   #r := FALSE;
   #a1 := W#16#0000;
   #a2 := W#16#0000;
   #activeDataBlock := 0;
   // PB17, STEP 5 network 1
   #r := ((NOT "ROLL_State".M[70, 1]) AND "ROLL_State".M[3, 3]);
   "ROLL_State".M[70, 0] := #r;
   // PB17, STEP 5 network 2
   #r := "ROLL_State".M[70, 0];
   IF #r THEN
       "ROLL_State".M[70, 1] := TRUE;
   END_IF;
   #r := "ROLL_IO".Input[0, 2];
   IF #r THEN
       "ROLL_State".M[70, 1] := FALSE;
   END_IF;
   // PB17, STEP 5 network 3
   #r := ((("ROLL_IO".Input[0, 1] AND "ROLL_State".M[74, 1]) OR ("ROLL_IO".Input[0, 2] AND "ROLL_State".M[64, 0])) AND "ROLL_State".M[29, 1]);
   "ROLL_IO".Output[112, 0] := #r;
   // PB17, STEP 5 network 4
   #r := ((("ROLL_IO".Input[0, 1] AND "ROLL_State".M[74, 5]) OR ("ROLL_IO".Input[0, 2] AND "ROLL_State".M[64, 1])) AND "ROLL_State".M[29, 1]);
   "ROLL_IO".Output[112, 5] := #r;
   // PB17, STEP 5 network 5
   #r := (((("ROLL_IO".Input[0, 1] AND "ROLL_State".M[78, 4]) OR ("ROLL_IO".Input[0, 2] AND "ROLL_State".M[64, 4])) AND "ROLL_State".M[29, 0]) OR ("ROLL_IO".Output[113, 1] AND "ROLL_IO".Output[113, 3]));
   "ROLL_IO".Output[113, 1] := #r;
   // PB17, STEP 5 network 6
   #r := (((NOT "ROLL_State".M[71, 4]) AND "ROLL_State".M[71, 3]) OR ((("ROLL_IO".Input[0, 1] AND "ROLL_State".M[78, 6]) OR ("ROLL_IO".Input[0, 2] AND "ROLL_State".M[64, 5])) AND "ROLL_State".M[29, 0]));
   "ROLL_State".M[71, 3] := #r;
   // PB17, STEP 5 network 7
   #r := "ROLL_State".M[71, 3];
   "ROLL_IO".Output[113, 3] := #r;
   // PB17, STEP 5 network 8
   #r := (((NOT "ROLL_State".M[71, 3]) AND "ROLL_State".M[71, 4]) OR ((((NOT "ROLL_State".M[64, 5]) AND ((NOT "ROLL_State".M[20, 2]) OR "ROLL_IO".Input[124, 5]) AND "ROLL_IO".Input[0, 2]) OR ("ROLL_IO".Input[0, 1] AND "ROLL_State".M[78, 7])) AND "ROLL_State".M[29, 0]));
   "ROLL_State".M[71, 4] := #r;
   // PB17, STEP 5 network 9
   #r := "ROLL_State".M[71, 4];
   "ROLL_IO".Output[113, 2] := #r;
   // PB17, STEP 5 network 10
   #r := (("ROLL_IO".Input[0, 1] AND "ROLL_State".M[75, 4]) OR ("ROLL_IO".Input[0, 2] AND "ROLL_State".M[35, 2] AND "ROLL_State".M[65, 0]));
   "ROLL_State".M[79, 5] := #r;
   // PB17, STEP 5 network 11
   #r := ((NOT "ROLL_IO".Output[23, 0]) AND (NOT "ROLL_IO".Output[23, 4]) AND (NOT "ROLL_State".M[10, 3]) AND (NOT "ROLL_State".M[5, 0]) AND ((NOT "ROLL_IO".Input[11, 4]) OR (NOT "ROLL_IO".Input[11, 6])) AND "ROLL_IO".Input[11, 7] AND "ROLL_IO".Input[12, 5] AND "ROLL_IO".Input[12, 7] AND "ROLL_IO".Input[14, 0] AND "ROLL_State".M[29, 0] AND "ROLL_State".M[79, 5]);
   "ROLL_IO".Output[23, 1] := #r;
   // PB17, STEP 5 network 12
   #r := (("ROLL_IO".Input[0, 1] AND "ROLL_State".M[75, 5]) OR ("ROLL_IO".Input[0, 2] AND "ROLL_State".M[35, 2] AND "ROLL_State".M[65, 5]));
   "ROLL_State".M[79, 6] := #r;
   // PB17, STEP 5 network 13
   #r := ((NOT "ROLL_IO".Output[23, 1]) AND (NOT "ROLL_IO".Output[23, 4]) AND (NOT "ROLL_State".M[10, 2]) AND (NOT "ROLL_State".M[5, 0]) AND (((NOT "ROLL_IO".Input[119, 0]) AND "ROLL_State".M[0, 3]) OR (NOT "ROLL_IO".Input[11, 0]) OR (NOT "ROLL_IO".Input[11, 6])) AND "ROLL_IO".Input[11, 7] AND "ROLL_IO".Input[12, 5] AND "ROLL_IO".Input[12, 7] AND "ROLL_IO".Input[14, 0] AND "ROLL_State".M[29, 0] AND "ROLL_State".M[79, 6]);
   "ROLL_IO".Output[23, 0] := #r;
   // PB17, STEP 5 network 14
   #r := ((("ROLL_IO".Input[0, 1] AND "ROLL_State".M[75, 6]) OR ("ROLL_IO".Input[0, 2] AND "ROLL_State".M[35, 2] AND "ROLL_State".M[65, 6])) AND ("ROLL_IO".Output[23, 0] OR "ROLL_IO".Output[23, 1]));
   "ROLL_IO".Output[23, 3] := #r;
   // PB17, STEP 5 network 15
   #r := ((NOT "ROLL_IO".Output[23, 3]) AND ("ROLL_IO".Output[23, 0] OR "ROLL_IO".Output[23, 1]) AND ("ROLL_IO".Input[0, 1] OR "ROLL_State".M[31, 5]) AND "ROLL_State".M[29, 0]);
   "ROLL_IO".Output[23, 2] := #r;
   // PB17, STEP 5 network 16
   #r := (("ROLL_IO".Input[0, 1] AND "ROLL_State".M[76, 2]) OR ("ROLL_IO".Input[0, 2] AND "ROLL_State".M[35, 2] AND "ROLL_State".M[66, 4]));
   "ROLL_State".M[80, 0] := #r;
   // PB17, STEP 5 network 17
   #r := ((NOT "ROLL_IO".Output[23, 4]) AND (NOT "ROLL_State".M[10, 1]) AND (NOT "ROLL_State".M[5, 2]) AND (NOT "ROLL_State".M[9, 0]) AND ((NOT "ROLL_IO".Input[12, 5]) OR (NOT "ROLL_IO".Input[12, 7])) AND ("ROLL_IO".Input[124, 2] OR "ROLL_State".M[0, 4]) AND "ROLL_IO".Input[13, 0] AND "ROLL_IO".Input[13, 7] AND "ROLL_IO".Input[14, 0] AND "ROLL_State".M[29, 0] AND "ROLL_State".M[80, 0]);
   "ROLL_IO".Output[23, 5] := #r;
   // PB17, STEP 5 network 18
   #r := (("ROLL_IO".Input[0, 1] AND "ROLL_State".M[77, 0]) OR ("ROLL_IO".Input[0, 2] AND "ROLL_State".M[35, 2] AND "ROLL_State".M[66, 7]));
   "ROLL_State".M[80, 1] := #r;
   // PB17, STEP 5 network 19
   #r := "ROLL_IO".Input[12, 5];
   IF #r THEN
       "ROLL_State".M[80, 2] := TRUE;
   END_IF;
   #r := "ROLL_IO".Input[12, 1];
   IF #r THEN
       "ROLL_State".M[80, 2] := FALSE;
   END_IF;
   // PB17, STEP 5 network 20
   #r := (((("ROLL_IO".Input[11, 1] OR "ROLL_IO".Input[11, 2] OR "ROLL_IO".Input[11, 3] OR "ROLL_IO".Input[11, 4] OR "ROLL_IO".Input[119, 6] OR "ROLL_IO".Input[119, 7] OR "ROLL_IO".Input[120, 0] OR "ROLL_IO".Input[120, 1]) AND "ROLL_IO".Input[12, 1]) OR ("ROLL_IO".Input[11, 0] AND "ROLL_IO".Input[12, 1])) AND "ROLL_IO".Input[12, 7]);
   "ROLL_State".M[80, 6] := #r;
   // PB17, STEP 5 network 21
   #r := (("ROLL_IO".Input[11, 0] OR "ROLL_IO".Input[11, 1] OR "ROLL_IO".Input[11, 2] OR "ROLL_IO".Input[11, 3] OR "ROLL_IO".Input[11, 4] OR "ROLL_IO".Input[119, 6] OR "ROLL_IO".Input[119, 7] OR "ROLL_IO".Input[120, 0] OR "ROLL_IO".Input[120, 1]) AND "ROLL_IO".Input[12, 5] AND "ROLL_IO".Input[12, 7]);
   "ROLL_State".M[80, 7] := #r;
   // PB17, STEP 5 network 22
   #r := ((NOT "ROLL_IO".Output[23, 0]) AND (NOT "ROLL_IO".Output[23, 1]) AND (NOT "ROLL_IO".Output[23, 5]) AND (NOT "ROLL_State".M[10, 0]) AND (NOT "ROLL_State".M[5, 2]) AND (NOT "ROLL_State".M[80, 6]) AND ("ROLL_IO".Input[124, 2] OR "ROLL_State".M[0, 4]) AND "ROLL_IO".Input[13, 0] AND "ROLL_IO".Input[14, 0] AND "ROLL_State".M[29, 0] AND "ROLL_State".M[80, 1]);
   "ROLL_IO".Output[23, 4] := #r;
   // PB17, STEP 5 network 23
   #r := ((NOT "ROLL_State".M[68, 2]) AND (((NOT "ROLL_IO".Input[12, 5]) AND "ROLL_IO".Output[23, 5]) OR ("ROLL_IO".Output[23, 4] AND "ROLL_State".M[80, 2])));
   "ROLL_IO".Output[23, 7] := #r;
   // PB17, STEP 5 network 24
   #r := ((NOT "ROLL_IO".Output[23, 7]) AND ("ROLL_IO".Output[23, 4] OR "ROLL_IO".Output[23, 5]));
   "ROLL_IO".Output[23, 6] := #r;
   // PB17, STEP 5 network 25
   #r := (("ROLL_IO".Input[0, 1] AND "ROLL_State".M[77, 6]) OR ("ROLL_IO".Input[0, 2] AND "ROLL_State".M[35, 2] AND "ROLL_State".M[67, 0]));
   "ROLL_State".M[80, 3] := #r;
   // PB17, STEP 5 network 26
   #r := ((NOT "ROLL_IO".Output[112, 1]) AND (NOT "ROLL_IO".Output[113, 3]) AND (NOT "ROLL_IO".Input[124, 2]) AND (NOT "ROLL_State".M[10, 5]) AND (NOT "ROLL_State".M[70, 2]) AND (NOT "ROLL_State".M[9, 3]) AND "ROLL_IO".Input[11, 0] AND "ROLL_IO".Input[11, 6] AND "ROLL_IO".Input[12, 1] AND "ROLL_IO".Input[12, 7] AND "ROLL_State".M[29, 0] AND "ROLL_State".M[80, 3]);
   "ROLL_IO".Output[112, 2] := #r;
   // PB17, STEP 5 network 27
   #r := (("ROLL_IO".Input[0, 1] AND "ROLL_State".M[77, 4]) OR ("ROLL_IO".Input[0, 2] AND "ROLL_State".M[35, 2] AND "ROLL_State".M[67, 1]));
   "ROLL_State".M[80, 4] := #r;
   // PB17, STEP 5 network 28
   #r := ((NOT "ROLL_IO".Output[112, 2]) AND (NOT "ROLL_IO".Output[113, 3]) AND (NOT "ROLL_IO".Input[124, 1]) AND (NOT "ROLL_State".M[10, 4]) AND (NOT "ROLL_State".M[70, 2]) AND (NOT "ROLL_State".M[70, 3]) AND (NOT "ROLL_State".M[9, 3]) AND "ROLL_IO".Input[11, 0] AND "ROLL_IO".Input[11, 6] AND "ROLL_IO".Input[12, 1] AND "ROLL_IO".Input[12, 7] AND "ROLL_State".M[29, 0] AND "ROLL_State".M[80, 4]);
   "ROLL_IO".Output[112, 1] := #r;
   // PB17, STEP 5 network 29
   #r := ((("ROLL_IO".Input[0, 1] AND "ROLL_State".M[77, 7]) OR ("ROLL_IO".Input[0, 2] AND "ROLL_State".M[35, 2] AND "ROLL_State".M[67, 5])) AND "ROLL_State".M[29, 0]);
   "ROLL_IO".Output[112, 4] := #r;
   // PB17, STEP 5 network 30
   #r := ((("ROLL_IO".Input[0, 1] AND "ROLL_State".M[78, 0]) OR ("ROLL_IO".Input[0, 2] AND "ROLL_State".M[35, 2] AND "ROLL_State".M[67, 6])) AND "ROLL_State".M[29, 0]);
   "ROLL_IO".Output[112, 3] := #r;
   // PB17, STEP 5 network 31
   #r := ((NOT "ROLL_State".M[16, 0]) AND (NOT "ROLL_State".M[16, 1]) AND (NOT "ROLL_State".M[16, 2]) AND (NOT "ROLL_State".M[16, 4]) AND "ROLL_State".M[37, 2]);
   "ROLL_State".M[81, 4] := #r;
   // PB17, STEP 5 network 32
   RETURN;
END_FUNCTION

FUNCTION "ROLL_PB18" : Void   // FC26, SCL
{ S7_Optimized_Access := 'TRUE' }
VERSION : 0.1
// stored: AutoNumber true, IsIECCheckEnabled false, SetENOAutomatically false, UDAEnableTagReadback false
   VAR_TEMP
      r : Bool;
      a1 : Word;
      a2 : Word;
      activeDataBlock : Int;
      comparisonResults : Array[0..0] of Bool;
   END_VAR
BEGIN

   #r := FALSE;
   #a1 := W#16#0000;
   #a2 := W#16#0000;
   #activeDataBlock := 0;
   // PB18, STEP 5 network 1
   #r := ("ROLL_State".M[70, 2] OR "ROLL_State".M[70, 3] OR "ROLL_State".M[70, 4] OR "ROLL_State".M[70, 6] OR "ROLL_State".M[71, 0]);
   "ROLL_State".M[80, 5] := #r;
   // PB18, STEP 5 network 2
   #r := (((NOT "ROLL_IO".Output[112, 0]) AND (NOT "ROLL_IO".Output[112, 5]) AND "ROLL_State".M[20, 5]) OR ((NOT "ROLL_IO".Output[112, 0]) AND "ROLL_State".M[20, 3]) OR ((NOT "ROLL_IO".Output[112, 5]) AND "ROLL_State".M[20, 4]) OR ((NOT "ROLL_IO".Output[17, 7]) AND "ROLL_State".M[20, 7]) OR (("ROLL_State".M[20, 1] OR "ROLL_State".M[20, 2]) AND "ROLL_State".M[28, 4]));
   "ROLL_State".M[250, 0] := #r;
   // PB18, STEP 5 network 3
   #r := (((NOT "ROLL_IO".Output[113, 0]) AND "ROLL_State".M[22, 2]) OR ((NOT "ROLL_IO".Output[113, 1]) AND "ROLL_State".M[22, 3]) OR ((NOT "ROLL_IO".Output[113, 3]) AND "ROLL_IO".Output[113, 2] AND "ROLL_State".M[22, 4]) OR ((NOT "ROLL_IO".Output[113, 5]) AND "ROLL_IO".Output[113, 4] AND "ROLL_State".M[22, 5]) OR ("ROLL_IO".Input[124, 1] AND "ROLL_State".M[22, 0]) OR ("ROLL_IO".Input[124, 4] AND "ROLL_State".M[22, 1]) OR "ROLL_State".M[250, 0]);
   "ROLL_State".M[250, 0] := #r;
   // PB18, STEP 5 network 4
   #r := ((("ROLL_IO".Input[11, 1] OR "ROLL_IO".Input[11, 2] OR "ROLL_IO".Input[11, 3] OR "ROLL_IO".Input[11, 4] OR "ROLL_IO".Input[119, 6] OR "ROLL_IO".Input[119, 7] OR "ROLL_IO".Input[120, 0] OR "ROLL_IO".Input[120, 1]) AND "ROLL_IO".Input[12, 5] AND "ROLL_IO".Input[12, 7] AND "ROLL_State".M[23, 0]) OR (("ROLL_State".M[23, 2] OR "ROLL_State".M[23, 3]) AND "ROLL_State".M[63, 1]) OR ("ROLL_IO".Input[11, 0] AND "ROLL_IO".Input[11, 6] AND "ROLL_State".M[23, 1]) OR ("ROLL_IO".Input[11, 0] AND "ROLL_IO".Input[12, 1] AND "ROLL_IO".Input[12, 7] AND "ROLL_State".M[23, 0]) OR "ROLL_State".M[250, 0]);
   "ROLL_State".M[250, 0] := #r;
   // PB18, STEP 5 network 5
   #r := (((NOT "ROLL_IO".Output[20, 1]) AND "ROLL_State".M[24, 1]) OR "ROLL_State".M[250, 0]);
   "ROLL_State".M[250, 0] := #r;
   // PB18, STEP 5 network 6
   #r := ((((NOT "ROLL_IO".Output[20, 4]) OR (NOT "ROLL_IO".Output[22, 6])) AND "ROLL_State".M[25, 0]) OR "ROLL_State".M[250, 0]);
   "ROLL_State".M[250, 0] := #r;
   // PB18, STEP 5 network 7
   #r := (((NOT "ROLL_IO".Output[20, 5]) AND "ROLL_State".M[26, 6]) OR ((NOT "ROLL_IO".Output[20, 6]) AND "ROLL_State".M[26, 0]) OR ((NOT "ROLL_IO".Output[21, 4]) AND "ROLL_State".M[26, 5]) OR "ROLL_State".M[250, 0]);
   "ROLL_State".M[250, 0] := #r;
   // PB18, STEP 5 network 8
   #r := (((NOT "ROLL_IO".Output[20, 6]) AND "ROLL_State".M[27, 4]) OR ((NOT "ROLL_IO".Output[21, 6]) AND "ROLL_State".M[27, 5]) OR ((NOT "ROLL_State".M[80, 5]) AND "ROLL_State".M[27, 7]) OR "ROLL_State".M[250, 0]);
   "ROLL_State".M[250, 0] := #r;
   // PB18, STEP 5 network 9
   #r := ((("ROLL_IO".Output[112, 0] OR "ROLL_IO".Output[112, 5]) AND "ROLL_State".M[20, 5]) OR ("ROLL_IO".Output[112, 0] AND "ROLL_State".M[20, 3]) OR ("ROLL_IO".Output[112, 5] AND "ROLL_State".M[20, 4]) OR ("ROLL_IO".Output[17, 7] AND "ROLL_State".M[20, 7]));
   "ROLL_State".M[252, 0] := #r;
   // PB18, STEP 5 network 10
   #r := (((NOT "ROLL_IO".Output[113, 2]) AND "ROLL_IO".Output[113, 3] AND "ROLL_State".M[22, 4]) OR ((NOT "ROLL_IO".Output[113, 4]) AND "ROLL_IO".Output[113, 5] AND "ROLL_State".M[22, 5]) OR ("ROLL_IO".Output[113, 0] AND "ROLL_State".M[22, 2]) OR ("ROLL_IO".Output[113, 1] AND "ROLL_State".M[22, 3]) OR ("ROLL_IO".Input[124, 2] AND "ROLL_State".M[22, 0]) OR ("ROLL_IO".Input[124, 5] AND "ROLL_State".M[22, 1]) OR "ROLL_State".M[252, 0]);
   "ROLL_State".M[252, 0] := #r;
   // PB18, STEP 5 network 11
   #r := (((NOT "ROLL_IO".Output[23, 1]) AND ("ROLL_IO".Input[11, 1] OR "ROLL_IO".Input[11, 2] OR "ROLL_IO".Input[11, 3] OR "ROLL_IO".Input[11, 4] OR "ROLL_IO".Input[119, 6] OR "ROLL_IO".Input[119, 7] OR "ROLL_IO".Input[120, 0] OR "ROLL_IO".Input[120, 1]) AND "ROLL_IO".Input[11, 6] AND "ROLL_State".M[23, 1]) OR ((NOT "ROLL_State".M[63, 1]) AND ("ROLL_State".M[23, 2] OR "ROLL_State".M[23, 3])) OR (((("ROLL_IO".Input[11, 1] OR "ROLL_IO".Input[11, 2] OR "ROLL_IO".Input[11, 3] OR "ROLL_IO".Input[11, 4] OR "ROLL_IO".Input[119, 6] OR "ROLL_IO".Input[119, 7] OR "ROLL_IO".Input[120, 0] OR "ROLL_IO".Input[120, 1]) AND "ROLL_IO".Input[12, 1]) OR ("ROLL_IO".Input[11, 0] AND "ROLL_IO".Input[12, 5])) AND "ROLL_IO".Input[12, 7] AND "ROLL_State".M[23, 0]) OR "ROLL_State".M[252, 0]);
   "ROLL_State".M[252, 0] := #r;
   // PB18, STEP 5 network 12
   #r := (("ROLL_IO".Output[20, 1] AND "ROLL_State".M[24, 1]) OR "ROLL_State".M[252, 0]);
   "ROLL_State".M[252, 0] := #r;
   // PB18, STEP 5 network 13
   #r := (("ROLL_IO".Output[20, 4] AND "ROLL_IO".Output[22, 6] AND "ROLL_State".M[25, 0]) OR "ROLL_State".M[252, 0]);
   "ROLL_State".M[252, 0] := #r;
   // PB18, STEP 5 network 14
   #r := (("ROLL_IO".Output[20, 6] AND "ROLL_State".M[26, 0]) OR "ROLL_State".M[252, 0]);
   "ROLL_State".M[252, 0] := #r;
   // PB18, STEP 5 network 15
   #r := (("ROLL_IO".Output[20, 5] AND "ROLL_State".M[26, 6]) OR ("ROLL_IO".Output[20, 6] AND "ROLL_State".M[27, 4]) OR ("ROLL_IO".Output[21, 4] AND "ROLL_State".M[26, 5]) OR ("ROLL_IO".Output[21, 6] AND "ROLL_State".M[27, 5]) OR ("ROLL_State".M[27, 7] AND "ROLL_State".M[80, 5]) OR "ROLL_State".M[252, 0]);
   "ROLL_State".M[252, 0] := #r;
   // PB18, STEP 5 network 16
   RETURN;
END_FUNCTION

FUNCTION "ROLL_PB19" : Void   // FC27, SCL
{ S7_Optimized_Access := 'TRUE' }
VERSION : 0.1
// stored: AutoNumber true, IsIECCheckEnabled false, SetENOAutomatically false, UDAEnableTagReadback false
   VAR_TEMP
      r : Bool;
      a1 : Word;
      a2 : Word;
      activeDataBlock : Int;
      comparisonResults : Array[0..0] of Bool;
   END_VAR
BEGIN

   #r := FALSE;
   #a1 := W#16#0000;
   #a2 := W#16#0000;
   #activeDataBlock := 0;
   // PB19, STEP 5 network 1
   #r := ((NOT "ROLL_IO".Input[3, 6]) AND (NOT "ROLL_State".M[5, 6]) AND (NOT "ROLL_State".M[6, 0]) AND (NOT "ROLL_State".M[6, 2]) AND ("ROLL_IO".Input[3, 1] OR "ROLL_State".M[31, 5]) AND "ROLL_IO".Input[5, 2] AND "ROLL_IO".Input[5, 4] AND "ROLL_State".M[4, 1]);
   "ROLL_State".M[82, 0] := #r;
   // PB19, STEP 5 network 2
   #r := ((NOT "ROLL_IO".Input[3, 6]) AND (NOT "ROLL_State".M[12, 0]) AND (NOT "ROLL_State".M[5, 3]) AND (NOT "ROLL_State".M[5, 6]) AND ("ROLL_IO".Input[3, 1] OR "ROLL_State".M[31, 5]) AND "ROLL_IO".Input[8, 3] AND "ROLL_IO".Input[8, 5] AND "ROLL_State".M[4, 1]);
   "ROLL_State".M[82, 2] := #r;
   // PB19, STEP 5 network 3
   #r := ("ROLL_State".M[31, 5] AND "ROLL_State".M[40, 0]);
   IF #r THEN
       "ROLL_State".M[82, 3] := TRUE;
   END_IF;
   #r := (NOT "ROLL_State".M[31, 5]);
   IF #r THEN
       "ROLL_State".M[82, 3] := FALSE;
   END_IF;
   // PB19, STEP 5 network 4
   #r := ((NOT "ROLL_State".M[110, 1]) AND (NOT "ROLL_State".M[110, 2]) AND "ROLL_State".M[110, 0] AND "ROLL_State".M[110, 3] AND "ROLL_State".M[40, 0]);
   "ROLL_State".M[240, 0] := #r;
   // PB19, STEP 5 network 5
   #r := (((NOT "ROLL_State".M[110, 2]) AND "ROLL_State".M[110, 0] AND "ROLL_State".M[110, 1] AND "ROLL_State".M[110, 3] AND "ROLL_State".M[41, 1]) OR "ROLL_State".M[240, 0]);
   "ROLL_State".M[240, 0] := #r;
   // PB19, STEP 5 network 6
   #r := (((NOT "ROLL_State".M[110, 1]) AND "ROLL_State".M[110, 0] AND "ROLL_State".M[110, 2] AND "ROLL_State".M[110, 3] AND "ROLL_State".M[41, 1]) OR "ROLL_State".M[240, 0]);
   "ROLL_State".M[240, 0] := #r;
   // PB19, STEP 5 network 7
   #r := (("ROLL_State".M[110, 0] AND "ROLL_State".M[110, 1] AND "ROLL_State".M[110, 2] AND "ROLL_State".M[110, 3] AND "ROLL_State".M[41, 1]) OR "ROLL_State".M[240, 0]);
   "ROLL_State".M[240, 0] := #r;
   // PB19, STEP 5 network 8
   #r := ("ROLL_State".M[240, 0] AND "ROLL_State".M[31, 5]);
   IF #r THEN
       "ROLL_State".M[82, 4] := TRUE;
   END_IF;
   #r := ((NOT "ROLL_State".M[31, 5]) OR "ROLL_State".M[45, 5]);
   IF #r THEN
       "ROLL_State".M[82, 4] := FALSE;
   END_IF;
   // PB19, STEP 5 network 9
   #r := ((NOT "ROLL_IO".Output[17, 3]) AND (NOT "ROLL_State".M[82, 4]) AND (NOT "ROLL_State".S5Timers[91].Q) AND ("ROLL_State".M[82, 3] OR "ROLL_State".S5Timers[22].Q) AND "ROLL_IO".Input[8, 5]);
   "ROLL_IO".Output[17, 2] := #r;
   // PB19, STEP 5 network 10
   #r := ((NOT "ROLL_IO".Output[17, 2]) AND (NOT "ROLL_State".S5Timers[90].Q) AND "ROLL_IO".Input[3, 0] AND "ROLL_IO".Input[8, 5] AND "ROLL_State".M[82, 4]);
   "ROLL_IO".Output[17, 3] := #r;
   // PB19, STEP 5 network 11
   #a2 := #a1;
   #a1 := W#16#3060;
   #r := "ROLL_IO".Output[18, 0];
   "ROLL_TimerOp"(Number := 22,
                  Operation := 1,
                  Signal := #r,
                  Preset := #a1);
   // PB19, STEP 5 network 12
   #a2 := #a1;
   #a1 := W#16#1005;
   #r := "ROLL_IO".Output[17, 2];
   "ROLL_TimerOp"(Number := 90,
                  Operation := 1,
                  Signal := #r,
                  Preset := #a1);
   // PB19, STEP 5 network 13
   #a2 := #a1;
   #a1 := W#16#1040;
   #r := "ROLL_IO".Output[17, 3];
   "ROLL_TimerOp"(Number := 91,
                  Operation := 1,
                  Signal := #r,
                  Preset := #a1);
   // PB19, STEP 5 network 14
   #r := ((NOT "ROLL_State".M[12, 0]) AND (NOT "ROLL_State".M[19, 7]) AND ("ROLL_IO".Output[17, 2] OR "ROLL_IO".Output[17, 3] OR "ROLL_State".S5Timers[90].Q OR "ROLL_State".S5Timers[91].Q) AND ("ROLL_State".M[82, 3] OR "ROLL_State".M[82, 4]) AND "ROLL_IO".Input[8, 3] AND "ROLL_IO".Input[8, 4] AND "ROLL_State".M[82, 2]);
   "ROLL_IO".Output[18, 0] := #r;
   // PB19, STEP 5 network 15
   #r := "ROLL_IO".Output[18, 0];
   "ROLL_IO".Output[18, 1] := #r;
   // PB19, STEP 5 network 16
   #r := ("ROLL_IO".Output[18, 0] AND "ROLL_State".M[82, 4]);
   "ROLL_IO".Output[18, 2] := #r;
   // PB19, STEP 5 network 17
   #r := ("ROLL_IO".Output[18, 0] AND "ROLL_State".M[82, 4]);
   "ROLL_IO".Output[18, 3] := #r;
   // PB19, STEP 5 network 18
   RETURN;
END_FUNCTION

FUNCTION "ROLL_PB2" : Void   // FC14, SCL
{ S7_Optimized_Access := 'TRUE' }
VERSION : 0.1
// stored: AutoNumber true, IsIECCheckEnabled false, SetENOAutomatically false, UDAEnableTagReadback false
   VAR_TEMP
      r : Bool;
      a1 : Word;
      a2 : Word;
      activeDataBlock : Int;
      comparisonResults : Array[0..0] of Bool;
   END_VAR
BEGIN

   #r := FALSE;
   #a1 := W#16#0000;
   #a2 := W#16#0000;
   #activeDataBlock := 0;
   // PB2, STEP 5 network 1
   #r := ((NOT "ROLL_State".M[0, 1]) AND "ROLL_State".S5Timers[11].Q);
   "ROLL_State".M[4, 1] := #r;
   // PB2, STEP 5 network 2
   #r := ((NOT "ROLL_State".M[4, 1]) OR "ROLL_IO".Input[1, 0]);
   "ROLL_State".M[3, 1] := #r;
   // PB2, STEP 5 network 3
   #r := ((((NOT "ROLL_State".M[31, 4]) AND "ROLL_IO".Input[0, 4] AND "ROLL_State".M[4, 1]) OR "ROLL_State".M[31, 5]) AND "ROLL_IO".Input[0, 2]);
   "ROLL_State".M[4, 4] := #r;
   // PB2, STEP 5 network 4
   #r := (NOT "ROLL_IO".Input[11, 7]);
   IF #r THEN
       "ROLL_State".M[5, 0] := TRUE;
   END_IF;
   #r := "ROLL_State".M[3, 1];
   IF #r THEN
       "ROLL_State".M[5, 0] := FALSE;
   END_IF;
   // PB2, STEP 5 network 5
   #r := (NOT "ROLL_IO".Input[13, 5]);
   IF #r THEN
       "ROLL_State".M[5, 1] := TRUE;
   END_IF;
   #r := "ROLL_State".M[3, 1];
   IF #r THEN
       "ROLL_State".M[5, 1] := FALSE;
   END_IF;
   // PB2, STEP 5 network 6
   #r := (NOT "ROLL_IO".Input[13, 0]);
   IF #r THEN
       "ROLL_State".M[5, 2] := TRUE;
   END_IF;
   #r := "ROLL_State".M[3, 1];
   IF #r THEN
       "ROLL_State".M[5, 2] := FALSE;
   END_IF;
   // PB2, STEP 5 network 7
   #r := (NOT "ROLL_IO".Input[8, 5]);
   IF #r THEN
       "ROLL_State".M[5, 3] := TRUE;
   END_IF;
   #r := "ROLL_State".M[3, 1];
   IF #r THEN
       "ROLL_State".M[5, 3] := FALSE;
   END_IF;
   // PB2, STEP 5 network 8
   #r := "ROLL_State".M[0, 3];
   IF #r THEN
       "ROLL_State".M[5, 4] := TRUE;
   END_IF;
   #r := "ROLL_State".M[3, 1];
   IF #r THEN
       "ROLL_State".M[5, 4] := FALSE;
   END_IF;
   // PB2, STEP 5 network 9
   #r := "ROLL_State".M[0, 3];
   IF #r THEN
       "ROLL_State".M[5, 5] := TRUE;
   END_IF;
   #r := "ROLL_State".M[3, 1];
   IF #r THEN
       "ROLL_State".M[5, 5] := FALSE;
   END_IF;
   // PB2, STEP 5 network 10
   #r := "ROLL_IO".Input[3, 6];
   IF #r THEN
       "ROLL_State".M[5, 6] := TRUE;
   END_IF;
   #r := "ROLL_State".M[3, 1];
   IF #r THEN
       "ROLL_State".M[5, 6] := FALSE;
   END_IF;
   // PB2, STEP 5 network 11
   #r := (NOT "ROLL_IO".Input[3, 7]);
   IF #r THEN
       "ROLL_State".M[5, 7] := TRUE;
   END_IF;
   #r := "ROLL_State".M[3, 1];
   IF #r THEN
       "ROLL_State".M[5, 7] := FALSE;
   END_IF;
   // PB2, STEP 5 network 12
   #r := (NOT "ROLL_IO".Input[5, 2]);
   IF #r THEN
       "ROLL_State".M[6, 0] := TRUE;
   END_IF;
   #r := ("ROLL_IO".Input[5, 2] AND "ROLL_State".M[3, 1]);
   IF #r THEN
       "ROLL_State".M[6, 0] := FALSE;
   END_IF;
   // PB2, STEP 5 network 13
   #r := ((NOT "ROLL_IO".Input[5, 3]) AND "ROLL_State".S5Timers[31].Q);
   IF #r THEN
       "ROLL_State".M[6, 1] := TRUE;
   END_IF;
   #r := "ROLL_State".M[3, 1];
   IF #r THEN
       "ROLL_State".M[6, 1] := FALSE;
   END_IF;
   // PB2, STEP 5 network 14
   #r := (NOT "ROLL_IO".Input[5, 4]);
   IF #r THEN
       "ROLL_State".M[6, 2] := TRUE;
   END_IF;
   #r := ("ROLL_IO".Input[5, 4] AND "ROLL_State".M[3, 1]);
   IF #r THEN
       "ROLL_State".M[6, 2] := FALSE;
   END_IF;
   // PB2, STEP 5 network 15
   #r := ((NOT "ROLL_IO".Input[5, 5]) AND "ROLL_State".M[40, 5] AND "ROLL_State".S5Timers[17].Q);
   IF #r THEN
       "ROLL_State".M[6, 3] := TRUE;
   END_IF;
   #r := "ROLL_State".M[3, 1];
   IF #r THEN
       "ROLL_State".M[6, 3] := FALSE;
   END_IF;
   // PB2, STEP 5 network 16
   #r := ((NOT "ROLL_IO".Input[6, 0]) AND "ROLL_State".S5Timers[32].Q);
   IF #r THEN
       "ROLL_State".M[6, 4] := TRUE;
   END_IF;
   #r := "ROLL_State".M[3, 1];
   IF #r THEN
       "ROLL_State".M[6, 4] := FALSE;
   END_IF;
   // PB2, STEP 5 network 17
   #r := ((NOT "ROLL_IO".Input[6, 2]) AND "ROLL_State".S5Timers[33].Q);
   IF #r THEN
       "ROLL_State".M[6, 5] := TRUE;
   END_IF;
   #r := "ROLL_State".M[3, 1];
   IF #r THEN
       "ROLL_State".M[6, 5] := FALSE;
   END_IF;
   // PB2, STEP 5 network 18
   #r := "ROLL_State".M[0, 3];
   IF #r THEN
       "ROLL_State".M[6, 6] := TRUE;
   END_IF;
   #r := "ROLL_State".M[3, 1];
   IF #r THEN
       "ROLL_State".M[6, 6] := FALSE;
   END_IF;
   // PB2, STEP 5 network 19
   #r := ((NOT "ROLL_State".M[0, 3]) AND "ROLL_State".S5Timers[35].Q);
   IF #r THEN
       "ROLL_State".M[6, 7] := TRUE;
   END_IF;
   #r := "ROLL_State".M[3, 1];
   IF #r THEN
       "ROLL_State".M[6, 7] := FALSE;
   END_IF;
   // PB2, STEP 5 network 20
   #r := ((NOT "ROLL_State".M[0, 3]) AND "ROLL_State".S5Timers[36].Q);
   IF #r THEN
       "ROLL_State".M[7, 0] := TRUE;
   END_IF;
   #r := "ROLL_State".M[3, 1];
   IF #r THEN
       "ROLL_State".M[7, 0] := FALSE;
   END_IF;
   // PB2, STEP 5 network 21
   #r := ((NOT "ROLL_State".M[0, 3]) AND "ROLL_State".M[48, 1] AND "ROLL_State".S5Timers[37].Q);
   IF #r THEN
       "ROLL_State".M[7, 1] := TRUE;
   END_IF;
   #r := "ROLL_State".M[3, 1];
   IF #r THEN
       "ROLL_State".M[7, 1] := FALSE;
   END_IF;
   // PB2, STEP 5 network 22
   #r := ((NOT "ROLL_State".M[0, 3]) AND "ROLL_State".S5Timers[38].Q);
   IF #r THEN
       "ROLL_State".M[7, 2] := TRUE;
   END_IF;
   #r := "ROLL_State".M[3, 1];
   IF #r THEN
       "ROLL_State".M[7, 2] := FALSE;
   END_IF;
   // PB2, STEP 5 network 23
   #r := ((NOT "ROLL_IO".Input[5, 6]) AND "ROLL_State".S5Timers[16].Q);
   IF #r THEN
       "ROLL_State".M[7, 3] := TRUE;
   END_IF;
   #r := ("ROLL_IO".Input[5, 6] AND "ROLL_State".M[3, 1]);
   IF #r THEN
       "ROLL_State".M[7, 3] := FALSE;
   END_IF;
   // PB2, STEP 5 network 24
   #r := "ROLL_State".M[0, 3];
   IF #r THEN
       "ROLL_State".M[7, 4] := TRUE;
   END_IF;
   #r := "ROLL_State".M[3, 1];
   IF #r THEN
       "ROLL_State".M[7, 4] := FALSE;
   END_IF;
   // PB2, STEP 5 network 25
   #r := "ROLL_State".M[0, 3];
   IF #r THEN
       "ROLL_State".M[7, 5] := TRUE;
   END_IF;
   #r := "ROLL_State".M[3, 1];
   IF #r THEN
       "ROLL_State".M[7, 5] := FALSE;
   END_IF;
   // PB2, STEP 5 network 26
   #r := "ROLL_State".M[0, 3];
   IF #r THEN
       "ROLL_State".M[7, 6] := TRUE;
   END_IF;
   #r := "ROLL_State".M[3, 1];
   IF #r THEN
       "ROLL_State".M[7, 6] := FALSE;
   END_IF;
   // PB2, STEP 5 network 27
   #r := (NOT "ROLL_IO".Input[6, 7]);
   IF #r THEN
       "ROLL_State".M[7, 7] := TRUE;
   END_IF;
   #r := "ROLL_State".M[3, 1];
   IF #r THEN
       "ROLL_State".M[7, 7] := FALSE;
   END_IF;
   // PB2, STEP 5 network 28
   #a2 := #a1;
   #a1 := W#16#1050;
   #r := ((NOT "ROLL_IO".Input[7, 6]) AND "ROLL_IO".Output[20, 5]);
   "ROLL_TimerOp"(Number := 30,
                  Operation := 0,
                  Signal := #r,
                  Preset := #a1);
   #r := "ROLL_State".S5Timers[30].Q;
   IF #r THEN
       "ROLL_State".M[8, 6] := TRUE;
   END_IF;
   #r := "ROLL_State".M[3, 1];
   IF #r THEN
       "ROLL_State".M[8, 6] := FALSE;
   END_IF;
   // PB2, STEP 5 network 29
   #r := "ROLL_State".M[0, 3];
   IF #r THEN
       "ROLL_State".M[8, 7] := TRUE;
   END_IF;
   #r := "ROLL_State".M[3, 1];
   IF #r THEN
       "ROLL_State".M[8, 7] := FALSE;
   END_IF;
   // PB2, STEP 5 network 30
   #r := ((NOT "ROLL_IO".Input[13, 7]) AND "ROLL_State".M[4, 1]);
   IF #r THEN
       "ROLL_State".M[9, 0] := TRUE;
   END_IF;
   #r := ("ROLL_IO".Input[13, 7] AND "ROLL_State".M[3, 1]);
   IF #r THEN
       "ROLL_State".M[9, 0] := FALSE;
   END_IF;
   // PB2, STEP 5 network 31
   #r := "ROLL_State".M[0, 3];
   IF #r THEN
       "ROLL_State".M[9, 1] := TRUE;
   END_IF;
   #r := "ROLL_State".M[3, 1];
   IF #r THEN
       "ROLL_State".M[9, 1] := FALSE;
   END_IF;
   // PB2, STEP 5 network 32
   #r := ((NOT "ROLL_State".M[28, 4]) AND (NOT "ROLL_State".M[31, 5]) AND (((NOT "ROLL_State".M[20, 2]) AND ("ROLL_IO".Input[123, 5] OR "ROLL_IO".Input[123, 6])) OR "ROLL_State".M[70, 2] OR "ROLL_State".M[70, 3]) AND "ROLL_IO".Input[0, 4] AND "ROLL_State".M[4, 1]);
   IF #r THEN
       "ROLL_State".M[9, 2] := TRUE;
   END_IF;
   #r := "ROLL_State".M[3, 1];
   IF #r THEN
       "ROLL_State".M[9, 2] := FALSE;
   END_IF;
   // PB2, STEP 5 network 33
   #r := ("ROLL_State".M[4, 1] AND "ROLL_State".S5Timers[19].Q);
   IF #r THEN
       "ROLL_State".M[9, 3] := TRUE;
   END_IF;
   #r := "ROLL_State".M[3, 1];
   IF #r THEN
       "ROLL_State".M[9, 3] := FALSE;
   END_IF;
   // PB2, STEP 5 network 34
   #r := (((("ROLL_State".M[20, 4] OR "ROLL_State".M[20, 5]) AND "ROLL_IO".Input[0, 1] AND "ROLL_State".M[190, 6]) OR "ROLL_State".M[31, 5]) AND "ROLL_State".S5Timers[95].Q);
   "ROLL_State".M[9, 4] := #r;
   // PB2, STEP 5 network 35
   #r := "ROLL_State".M[0, 3];
   IF #r THEN
       "ROLL_State".M[9, 5] := TRUE;
   END_IF;
   #r := "ROLL_State".M[3, 1];
   IF #r THEN
       "ROLL_State".M[9, 5] := FALSE;
   END_IF;
   // PB2, STEP 5 network 36
   #r := "ROLL_State".M[0, 3];
   IF #r THEN
       "ROLL_State".M[9, 6] := TRUE;
   END_IF;
   #r := "ROLL_State".M[3, 1];
   IF #r THEN
       "ROLL_State".M[9, 6] := FALSE;
   END_IF;
   // PB2, STEP 5 network 37
   #r := "ROLL_State".M[0, 3];
   IF #r THEN
       "ROLL_State".M[9, 7] := TRUE;
   END_IF;
   #r := "ROLL_State".M[3, 1];
   IF #r THEN
       "ROLL_State".M[9, 7] := FALSE;
   END_IF;
   // PB2, STEP 5 network 38
   #r := ((NOT "ROLL_IO".Input[12, 0]) AND "ROLL_State".M[4, 1]);
   IF #r THEN
       "ROLL_State".M[10, 0] := TRUE;
   END_IF;
   #r := (((((NOT "ROLL_State".S5Timers[11].Q) AND "ROLL_IO".Input[3, 0]) OR "ROLL_IO".Input[12, 5]) AND "ROLL_State".M[3, 1]) OR (NOT "ROLL_State".M[4, 1]) OR "ROLL_State".M[0, 7]);
   IF #r THEN
       "ROLL_State".M[10, 0] := FALSE;
   END_IF;
   // PB2, STEP 5 network 39
   #r := ((NOT "ROLL_IO".Input[12, 6]) AND "ROLL_State".M[4, 1]);
   IF #r THEN
       "ROLL_State".M[10, 1] := TRUE;
   END_IF;
   #r := (((((NOT "ROLL_State".S5Timers[11].Q) AND "ROLL_IO".Input[3, 0]) OR "ROLL_IO".Input[12, 1]) AND "ROLL_State".M[3, 1]) OR (NOT "ROLL_State".M[4, 1]) OR "ROLL_State".M[0, 7]);
   IF #r THEN
       "ROLL_State".M[10, 1] := FALSE;
   END_IF;
   // PB2, STEP 5 network 40
   #r := "ROLL_State".M[0, 3];
   IF #r THEN
       "ROLL_State".M[10, 2] := TRUE;
   END_IF;
   #r := "ROLL_State".M[3, 1];
   IF #r THEN
       "ROLL_State".M[10, 2] := FALSE;
   END_IF;
   // PB2, STEP 5 network 41
   #r := "ROLL_State".M[0, 3];
   IF #r THEN
       "ROLL_State".M[10, 3] := TRUE;
   END_IF;
   #r := "ROLL_State".M[3, 1];
   IF #r THEN
       "ROLL_State".M[10, 3] := FALSE;
   END_IF;
   // PB2, STEP 5 network 42
   #r := "ROLL_State".M[0, 3];
   IF #r THEN
       "ROLL_State".M[10, 4] := TRUE;
   END_IF;
   #r := "ROLL_State".M[3, 1];
   IF #r THEN
       "ROLL_State".M[10, 4] := FALSE;
   END_IF;
   // PB2, STEP 5 network 43
   #r := "ROLL_State".M[0, 3];
   IF #r THEN
       "ROLL_State".M[10, 5] := TRUE;
   END_IF;
   #r := "ROLL_State".M[3, 1];
   IF #r THEN
       "ROLL_State".M[10, 5] := FALSE;
   END_IF;
   // PB2, STEP 5 network 44
   #r := "ROLL_State".M[0, 3];
   IF #r THEN
       "ROLL_State".M[10, 6] := TRUE;
   END_IF;
   #r := "ROLL_State".M[3, 1];
   IF #r THEN
       "ROLL_State".M[10, 6] := FALSE;
   END_IF;
   // PB2, STEP 5 network 45
   #r := "ROLL_State".M[0, 3];
   IF #r THEN
       "ROLL_State".M[10, 7] := TRUE;
   END_IF;
   #r := "ROLL_State".M[3, 1];
   IF #r THEN
       "ROLL_State".M[10, 7] := FALSE;
   END_IF;
   // PB2, STEP 5 network 46
   #r := ("ROLL_State".M[4, 1] AND "ROLL_State".M[63, 2]);
   IF #r THEN
       "ROLL_State".M[11, 0] := TRUE;
   END_IF;
   #r := "ROLL_State".M[3, 1];
   IF #r THEN
       "ROLL_State".M[11, 0] := FALSE;
   END_IF;
   // PB2, STEP 5 network 47
   #r := ("ROLL_IO".Input[13, 3] AND "ROLL_State".M[4, 1] AND "ROLL_State".S5Timers[112].Q);
   IF #r THEN
       "ROLL_State".M[11, 1] := TRUE;
   END_IF;
   #r := "ROLL_State".M[3, 1];
   IF #r THEN
       "ROLL_State".M[11, 1] := FALSE;
   END_IF;
   // PB2, STEP 5 network 48
   #r := ((NOT "ROLL_IO".Input[13, 3]) AND "ROLL_State".M[4, 1] AND "ROLL_State".S5Timers[15].Q);
   IF #r THEN
       "ROLL_State".M[11, 2] := TRUE;
   END_IF;
   #r := "ROLL_State".M[3, 1];
   IF #r THEN
       "ROLL_State".M[11, 2] := FALSE;
   END_IF;
   // PB2, STEP 5 network 49
   #r := ("ROLL_State".M[4, 1] AND "ROLL_State".M[63, 3]);
   IF #r THEN
       "ROLL_State".M[11, 3] := TRUE;
   END_IF;
   #r := "ROLL_State".M[3, 1];
   IF #r THEN
       "ROLL_State".M[11, 3] := FALSE;
   END_IF;
   // PB2, STEP 5 network 50
   #r := ("ROLL_State".M[190, 6] AND "ROLL_State".M[23, 2] AND "ROLL_State".M[60, 3]);
   IF #r THEN
       "ROLL_State".M[11, 4] := TRUE;
   END_IF;
   #r := "ROLL_State".M[3, 1];
   IF #r THEN
       "ROLL_State".M[11, 4] := FALSE;
   END_IF;
   // PB2, STEP 5 network 51
   #r := "ROLL_State".M[0, 3];
   IF #r THEN
       "ROLL_State".M[11, 5] := TRUE;
   END_IF;
   #r := "ROLL_State".M[3, 1];
   IF #r THEN
       "ROLL_State".M[11, 5] := FALSE;
   END_IF;
   // PB2, STEP 5 network 52
   #r := "ROLL_State".M[0, 3];
   IF #r THEN
       "ROLL_State".M[11, 6] := TRUE;
   END_IF;
   #r := "ROLL_State".M[3, 1];
   IF #r THEN
       "ROLL_State".M[11, 6] := FALSE;
   END_IF;
   // PB2, STEP 5 network 53
   #r := "ROLL_State".M[0, 3];
   IF #r THEN
       "ROLL_State".M[11, 7] := TRUE;
   END_IF;
   #r := "ROLL_State".M[3, 1];
   IF #r THEN
       "ROLL_State".M[11, 7] := FALSE;
   END_IF;
   // PB2, STEP 5 network 54
   #r := (NOT "ROLL_IO".Input[8, 3]);
   IF #r THEN
       "ROLL_State".M[12, 0] := TRUE;
   END_IF;
   #r := "ROLL_State".M[3, 1];
   IF #r THEN
       "ROLL_State".M[12, 0] := FALSE;
   END_IF;
   // PB2, STEP 5 network 55
   #r := ((NOT "ROLL_IO".Input[0, 7]) AND (NOT "ROLL_IO".Input[1, 4]) AND "ROLL_State".M[4, 4]);
   IF #r THEN
       "ROLL_State".M[12, 1] := TRUE;
   END_IF;
   #r := "ROLL_State".M[3, 1];
   IF #r THEN
       "ROLL_State".M[12, 1] := FALSE;
   END_IF;
   // PB2, STEP 5 network 56
   #r := "ROLL_State".M[0, 3];
   IF #r THEN
       "ROLL_State".M[12, 2] := TRUE;
   END_IF;
   #r := "ROLL_State".M[3, 1];
   IF #r THEN
       "ROLL_State".M[12, 2] := FALSE;
   END_IF;
   // PB2, STEP 5 network 57
   #r := "ROLL_State".M[0, 3];
   IF #r THEN
       "ROLL_State".M[12, 3] := TRUE;
   END_IF;
   #r := "ROLL_State".M[3, 1];
   IF #r THEN
       "ROLL_State".M[12, 3] := FALSE;
   END_IF;
   // PB2, STEP 5 network 58
   #r := "ROLL_State".M[0, 3];
   IF #r THEN
       "ROLL_State".M[13, 0] := TRUE;
   END_IF;
   #r := "ROLL_State".M[3, 1];
   IF #r THEN
       "ROLL_State".M[13, 0] := FALSE;
   END_IF;
   // PB2, STEP 5 network 59
   #r := (NOT "ROLL_IO".Input[3, 2]);
   IF #r THEN
       "ROLL_State".M[13, 1] := TRUE;
   END_IF;
   #r := "ROLL_State".M[3, 1];
   IF #r THEN
       "ROLL_State".M[13, 1] := FALSE;
   END_IF;
   // PB2, STEP 5 network 60
   #r := ((NOT "ROLL_IO".Input[4, 7]) AND "ROLL_IO".Input[0, 1] AND "ROLL_State".M[190, 6] AND "ROLL_State".M[27, 4]);
   IF #r THEN
       "ROLL_State".M[13, 2] := TRUE;
   END_IF;
   #r := "ROLL_State".M[3, 1];
   IF #r THEN
       "ROLL_State".M[13, 2] := FALSE;
   END_IF;
   // PB2, STEP 5 network 61
   #r := (NOT "ROLL_IO".Input[5, 0]);
   IF #r THEN
       "ROLL_State".M[13, 3] := TRUE;
   END_IF;
   #r := ("ROLL_IO".Input[5, 0] AND "ROLL_State".M[3, 1]);
   IF #r THEN
       "ROLL_State".M[13, 3] := FALSE;
   END_IF;
   // PB2, STEP 5 network 62
   #r := (NOT "ROLL_IO".Input[10, 7]);
   IF #r THEN
       "ROLL_State".M[13, 4] := TRUE;
   END_IF;
   #r := ("ROLL_IO".Input[10, 7] AND "ROLL_State".M[3, 1]);
   IF #r THEN
       "ROLL_State".M[13, 4] := FALSE;
   END_IF;
   // PB2, STEP 5 network 63
   #r := (NOT "ROLL_IO".Input[4, 5]);
   IF #r THEN
       "ROLL_State".M[13, 7] := TRUE;
   END_IF;
   #r := "ROLL_State".M[3, 1];
   IF #r THEN
       "ROLL_State".M[13, 7] := FALSE;
   END_IF;
   // PB2, STEP 5 network 64
   #a2 := #a1;
   #a1 := W#16#2020;
   #r := (((NOT "ROLL_IO".Input[10, 0]) OR (NOT "ROLL_IO".Input[10, 1]) OR (NOT "ROLL_IO".Input[10, 2]) OR (NOT "ROLL_IO".Input[10, 3])) AND "ROLL_IO".Output[19, 1]);
   "ROLL_TimerOp"(Number := 50,
                  Operation := 0,
                  Signal := #r,
                  Preset := #a1);
   // PB2, STEP 5 network 65
   #r := ((NOT "ROLL_IO".Input[10, 0]) AND "ROLL_State".S5Timers[50].Q);
   IF #r THEN
       "ROLL_State".M[14, 0] := TRUE;
   END_IF;
   #r := "ROLL_State".M[3, 1];
   IF #r THEN
       "ROLL_State".M[14, 0] := FALSE;
   END_IF;
   // PB2, STEP 5 network 66
   #r := ((NOT "ROLL_IO".Input[10, 1]) AND "ROLL_State".S5Timers[50].Q);
   IF #r THEN
       "ROLL_State".M[14, 1] := TRUE;
   END_IF;
   #r := "ROLL_State".M[3, 1];
   IF #r THEN
       "ROLL_State".M[14, 1] := FALSE;
   END_IF;
   // PB2, STEP 5 network 67
   #r := ((NOT "ROLL_IO".Input[10, 2]) AND "ROLL_State".S5Timers[50].Q);
   IF #r THEN
       "ROLL_State".M[14, 2] := TRUE;
   END_IF;
   #r := "ROLL_State".M[3, 1];
   IF #r THEN
       "ROLL_State".M[14, 2] := FALSE;
   END_IF;
   // PB2, STEP 5 network 68
   #r := ((NOT "ROLL_IO".Input[10, 3]) AND "ROLL_State".S5Timers[50].Q);
   IF #r THEN
       "ROLL_State".M[14, 3] := TRUE;
   END_IF;
   #r := "ROLL_State".M[3, 1];
   IF #r THEN
       "ROLL_State".M[14, 3] := FALSE;
   END_IF;
   // PB2, STEP 5 network 69
   #r := "ROLL_State".M[0, 3];
   IF #r THEN
       "ROLL_State".M[15, 2] := TRUE;
   END_IF;
   #r := "ROLL_State".M[3, 1];
   IF #r THEN
       "ROLL_State".M[15, 2] := FALSE;
   END_IF;
   // PB2, STEP 5 network 70
   #r := "ROLL_State".M[0, 3];
   IF #r THEN
       "ROLL_State".M[15, 3] := TRUE;
   END_IF;
   #r := "ROLL_State".M[3, 1];
   IF #r THEN
       "ROLL_State".M[15, 3] := FALSE;
   END_IF;
   // PB2, STEP 5 network 71
   #r := "ROLL_State".M[0, 3];
   IF #r THEN
       "ROLL_State".M[15, 4] := TRUE;
   END_IF;
   #r := "ROLL_State".M[3, 1];
   IF #r THEN
       "ROLL_State".M[15, 4] := FALSE;
   END_IF;
   // PB2, STEP 5 network 72
   #r := (NOT "ROLL_IO".Input[4, 0]);
   IF #r THEN
       "ROLL_State".M[15, 5] := TRUE;
   END_IF;
   #r := "ROLL_State".M[3, 1];
   IF #r THEN
       "ROLL_State".M[15, 5] := FALSE;
   END_IF;
   // PB2, STEP 5 network 73
   #r := (NOT "ROLL_IO".Input[4, 1]);
   IF #r THEN
       "ROLL_State".M[15, 6] := TRUE;
   END_IF;
   #r := "ROLL_State".M[3, 1];
   IF #r THEN
       "ROLL_State".M[15, 6] := FALSE;
   END_IF;
   // PB2, STEP 5 network 74
   #r := (NOT "ROLL_IO".Input[4, 2]);
   IF #r THEN
       "ROLL_State".M[15, 7] := TRUE;
   END_IF;
   #r := "ROLL_State".M[3, 1];
   IF #r THEN
       "ROLL_State".M[15, 7] := FALSE;
   END_IF;
   // PB2, STEP 5 network 75
   #r := "ROLL_State".M[16, 0];
   IF #r THEN
       "ROLL_State".M[16, 0] := TRUE;
   END_IF;
   #r := "ROLL_State".M[3, 1];
   IF #r THEN
       "ROLL_State".M[16, 0] := FALSE;
   END_IF;
   // PB2, STEP 5 network 76
   #r := "ROLL_State".M[16, 1];
   IF #r THEN
       "ROLL_State".M[16, 1] := TRUE;
   END_IF;
   #r := "ROLL_State".M[3, 1];
   IF #r THEN
       "ROLL_State".M[16, 1] := FALSE;
   END_IF;
   // PB2, STEP 5 network 77
   #r := "ROLL_State".M[16, 2];
   IF #r THEN
       "ROLL_State".M[16, 2] := TRUE;
   END_IF;
   #r := "ROLL_State".M[3, 1];
   IF #r THEN
       "ROLL_State".M[16, 2] := FALSE;
   END_IF;
   // PB2, STEP 5 network 78
   #r := ("ROLL_State".M[34, 1] AND "ROLL_State".M[4, 1]);
   IF #r THEN
       "ROLL_State".M[16, 3] := TRUE;
   END_IF;
   #r := "ROLL_State".M[3, 1];
   IF #r THEN
       "ROLL_State".M[16, 3] := FALSE;
   END_IF;
   // PB2, STEP 5 network 79
   #r := "ROLL_State".M[16, 4];
   IF #r THEN
       "ROLL_State".M[16, 4] := TRUE;
   END_IF;
   #r := ((NOT "ROLL_IO".Input[123, 1]) AND (NOT "ROLL_IO".Input[123, 4]) AND (NOT "ROLL_IO".Input[123, 5]) AND (NOT "ROLL_IO".Input[123, 6]) AND (NOT "ROLL_IO".Input[125, 0]) AND (NOT "ROLL_IO".Input[125, 1]) AND "ROLL_State".M[3, 1]);
   IF #r THEN
       "ROLL_State".M[16, 4] := FALSE;
   END_IF;
   // PB2, STEP 5 network 80
   #r := "ROLL_State".M[16, 5];
   IF #r THEN
       "ROLL_State".M[16, 5] := TRUE;
   END_IF;
   #r := "ROLL_State".M[3, 1];
   IF #r THEN
       "ROLL_State".M[16, 5] := FALSE;
   END_IF;
   // PB2, STEP 5 network 81
   #r := ((NOT "ROLL_IO".Input[3, 4]) AND "ROLL_State".M[4, 1]);
   IF #r THEN
       "ROLL_State".M[16, 6] := TRUE;
   END_IF;
   #r := ("ROLL_IO".Input[3, 4] AND "ROLL_State".M[3, 1]);
   IF #r THEN
       "ROLL_State".M[16, 6] := FALSE;
   END_IF;
   // PB2, STEP 5 network 82
   #r := ((NOT "ROLL_IO".Input[3, 1]) AND ((("ROLL_State".M[190, 5] OR "ROLL_State".M[190, 6]) AND "ROLL_IO".Input[0, 1]) OR "ROLL_State".M[4, 4]) AND "ROLL_State".M[4, 1]);
   IF #r THEN
       "ROLL_State".M[16, 7] := TRUE;
   END_IF;
   #r := "ROLL_State".M[3, 1];
   IF #r THEN
       "ROLL_State".M[16, 7] := FALSE;
   END_IF;
   // PB2, STEP 5 network 83
   #r := ((NOT "ROLL_IO".Input[3, 5]) AND "ROLL_State".M[4, 1]);
   IF #r THEN
       "ROLL_State".M[17, 0] := TRUE;
   END_IF;
   #r := ("ROLL_IO".Input[3, 5] AND "ROLL_State".M[3, 1]);
   IF #r THEN
       "ROLL_State".M[17, 0] := FALSE;
   END_IF;
   // PB2, STEP 5 network 84
   #r := "ROLL_State".M[0, 3];
   IF #r THEN
       "ROLL_State".M[17, 1] := TRUE;
   END_IF;
   #r := "ROLL_State".M[3, 1];
   IF #r THEN
       "ROLL_State".M[17, 1] := FALSE;
   END_IF;
   // PB2, STEP 5 network 85
   #r := "ROLL_State".M[0, 3];
   IF #r THEN
       "ROLL_State".M[17, 2] := TRUE;
   END_IF;
   #r := "ROLL_State".M[3, 1];
   IF #r THEN
       "ROLL_State".M[17, 2] := FALSE;
   END_IF;
   // PB2, STEP 5 network 86
   #r := "ROLL_State".M[0, 3];
   IF #r THEN
       "ROLL_State".M[17, 3] := TRUE;
   END_IF;
   #r := "ROLL_State".M[3, 1];
   IF #r THEN
       "ROLL_State".M[17, 3] := FALSE;
   END_IF;
   // PB2, STEP 5 network 87
   #r := "ROLL_State".M[0, 3];
   IF #r THEN
       "ROLL_State".M[17, 4] := TRUE;
   END_IF;
   #r := "ROLL_State".M[3, 1];
   IF #r THEN
       "ROLL_State".M[17, 4] := FALSE;
   END_IF;
   // PB2, STEP 5 network 88
   #r := "ROLL_State".M[0, 3];
   IF #r THEN
       "ROLL_State".M[17, 5] := TRUE;
   END_IF;
   #r := "ROLL_State".M[3, 1];
   IF #r THEN
       "ROLL_State".M[17, 5] := FALSE;
   END_IF;
   // PB2, STEP 5 network 89
   #r := "ROLL_State".M[0, 3];
   IF #r THEN
       "ROLL_State".M[17, 6] := TRUE;
   END_IF;
   #r := "ROLL_State".M[3, 1];
   IF #r THEN
       "ROLL_State".M[17, 6] := FALSE;
   END_IF;
   // PB2, STEP 5 network 90
   #r := "ROLL_State".M[0, 3];
   IF #r THEN
       "ROLL_State".M[17, 7] := TRUE;
   END_IF;
   #r := "ROLL_State".M[3, 1];
   IF #r THEN
       "ROLL_State".M[17, 7] := FALSE;
   END_IF;
   // PB2, STEP 5 network 91
   #r := "ROLL_State".M[0, 3];
   IF #r THEN
       "ROLL_State".M[18, 0] := TRUE;
   END_IF;
   #r := "ROLL_State".M[3, 1];
   IF #r THEN
       "ROLL_State".M[18, 0] := FALSE;
   END_IF;
   // PB2, STEP 5 network 92
   #r := ((NOT "ROLL_IO".Input[14, 0]) AND ((("ROLL_State".M[190, 5] OR "ROLL_State".M[190, 6]) AND ("ROLL_State".M[23, 0] OR "ROLL_State".M[23, 1] OR "ROLL_State".M[23, 2] OR "ROLL_State".M[23, 3])) OR ("ROLL_State".M[16, 3] AND "ROLL_State".M[31, 4] AND "ROLL_State".M[37, 2]) OR "ROLL_State".M[74, 0]));
   IF #r THEN
       "ROLL_State".M[18, 1] := TRUE;
   END_IF;
   #r := "ROLL_State".M[3, 1];
   IF #r THEN
       "ROLL_State".M[18, 1] := FALSE;
   END_IF;
   // PB2, STEP 5 network 93
   #r := "ROLL_State".M[0, 3];
   IF #r THEN
       "ROLL_State".M[18, 2] := TRUE;
   END_IF;
   #r := "ROLL_State".M[3, 1];
   IF #r THEN
       "ROLL_State".M[18, 2] := FALSE;
   END_IF;
   // PB2, STEP 5 network 94
   #r := "ROLL_State".M[0, 3];
   IF #r THEN
       "ROLL_State".M[18, 3] := TRUE;
   END_IF;
   #r := "ROLL_State".M[3, 1];
   IF #r THEN
       "ROLL_State".M[18, 3] := FALSE;
   END_IF;
   // PB2, STEP 5 network 95
   #r := "ROLL_State".M[0, 3];
   IF #r THEN
       "ROLL_State".M[18, 4] := TRUE;
   END_IF;
   #r := "ROLL_State".M[3, 1];
   IF #r THEN
       "ROLL_State".M[18, 4] := FALSE;
   END_IF;
   // PB2, STEP 5 network 96
   #r := "ROLL_State".M[0, 3];
   IF #r THEN
       "ROLL_State".M[18, 5] := TRUE;
   END_IF;
   #r := "ROLL_State".M[3, 1];
   IF #r THEN
       "ROLL_State".M[18, 5] := FALSE;
   END_IF;
   // PB2, STEP 5 network 97
   #r := "ROLL_State".M[0, 3];
   IF #r THEN
       "ROLL_State".M[18, 6] := TRUE;
   END_IF;
   #r := "ROLL_State".M[3, 1];
   IF #r THEN
       "ROLL_State".M[18, 6] := FALSE;
   END_IF;
   // PB2, STEP 5 network 98
   #r := "ROLL_State".M[0, 3];
   IF #r THEN
       "ROLL_State".M[18, 7] := TRUE;
   END_IF;
   #r := "ROLL_State".M[3, 1];
   IF #r THEN
       "ROLL_State".M[18, 7] := FALSE;
   END_IF;
   // PB2, STEP 5 network 99
   #r := "ROLL_State".M[0, 3];
   IF #r THEN
       "ROLL_State".M[19, 0] := TRUE;
   END_IF;
   #r := "ROLL_State".M[3, 1];
   IF #r THEN
       "ROLL_State".M[19, 0] := FALSE;
   END_IF;
   // PB2, STEP 5 network 100
   #r := "ROLL_State".M[0, 3];
   IF #r THEN
       "ROLL_State".M[19, 1] := TRUE;
   END_IF;
   #r := "ROLL_State".M[3, 1];
   IF #r THEN
       "ROLL_State".M[19, 1] := FALSE;
   END_IF;
   // PB2, STEP 5 network 101
   #r := "ROLL_State".M[0, 3];
   IF #r THEN
       "ROLL_State".M[19, 2] := TRUE;
   END_IF;
   #r := "ROLL_State".M[3, 1];
   IF #r THEN
       "ROLL_State".M[19, 2] := FALSE;
   END_IF;
   // PB2, STEP 5 network 102
   #r := "ROLL_State".M[0, 3];
   IF #r THEN
       "ROLL_State".M[19, 3] := TRUE;
   END_IF;
   #r := "ROLL_State".M[3, 1];
   IF #r THEN
       "ROLL_State".M[19, 3] := FALSE;
   END_IF;
   // PB2, STEP 5 network 103
   #r := "ROLL_State".M[0, 3];
   IF #r THEN
       "ROLL_State".M[19, 4] := TRUE;
   END_IF;
   #r := "ROLL_State".M[3, 1];
   IF #r THEN
       "ROLL_State".M[19, 4] := FALSE;
   END_IF;
   // PB2, STEP 5 network 104
   #r := "ROLL_State".M[0, 3];
   IF #r THEN
       "ROLL_State".M[19, 5] := TRUE;
   END_IF;
   #r := "ROLL_State".M[3, 1];
   IF #r THEN
       "ROLL_State".M[19, 5] := FALSE;
   END_IF;
   // PB2, STEP 5 network 105
   #r := "ROLL_State".M[0, 3];
   IF #r THEN
       "ROLL_State".M[19, 6] := TRUE;
   END_IF;
   #r := "ROLL_State".M[3, 1];
   IF #r THEN
       "ROLL_State".M[19, 6] := FALSE;
   END_IF;
   // PB2, STEP 5 network 106
   #r := "ROLL_State".M[0, 3];
   IF #r THEN
       "ROLL_State".M[19, 7] := TRUE;
   END_IF;
   #r := "ROLL_State".M[3, 1];
   IF #r THEN
       "ROLL_State".M[19, 7] := FALSE;
   END_IF;
   // PB2, STEP 5 network 107
   RETURN;
END_FUNCTION

FUNCTION "ROLL_PB20" : Void   // FC28, SCL
{ S7_Optimized_Access := 'TRUE' }
VERSION : 0.1
// stored: AutoNumber true, IsIECCheckEnabled false, SetENOAutomatically false, UDAEnableTagReadback false
   VAR_TEMP
      r : Bool;
      a1 : Word;
      a2 : Word;
      activeDataBlock : Int;
      comparisonResults : Array[0..0] of Bool;
   END_VAR
BEGIN

   #r := FALSE;
   #a1 := W#16#0000;
   #a2 := W#16#0000;
   #activeDataBlock := 0;
   // PB20, STEP 5 network 1
   #activeDataBlock := 15;
   // PB20, STEP 5 network 2
   #r := ((NOT "ROLL_IO".Input[7, 0]) AND (("ROLL_IO".Input[0, 1] AND "ROLL_State".M[190, 6] AND "ROLL_State".M[26, 5] AND "ROLL_State".M[4, 1]) OR ("ROLL_IO".Input[0, 2] AND "ROLL_State".M[0, 3])) AND "ROLL_State".M[4, 1]);
   "ROLL_State".M[8, 0] := #r;
   // PB20, STEP 5 network 3
   #r := ((NOT "ROLL_IO".Input[7, 1]) AND "ROLL_IO".Input[0, 2] AND "ROLL_IO".Input[1, 6] AND "ROLL_State".M[4, 1] AND "ROLL_State".S5Timers[61].Q);
   IF #r THEN
       "ROLL_State".M[8, 1] := TRUE;
   END_IF;
   #r := "ROLL_State".M[3, 1];
   IF #r THEN
       "ROLL_State".M[8, 1] := FALSE;
   END_IF;
   // PB20, STEP 5 network 4
   #a2 := #a1;
   #a1 := "ROLL_GetDW"(DbNumber := #activeDataBlock, Index := 61);
   #r := ((NOT "ROLL_IO".Input[7, 1]) AND "ROLL_IO".Input[0, 2] AND "ROLL_IO".Input[3, 1]);
   "ROLL_TimerOp"(Number := 61,
                  Operation := 0,
                  Signal := #r,
                  Preset := #a1);
   #r := ("ROLL_State".M[3, 1] AND "ROLL_State".M[4, 1]);
   "ROLL_TimerOp"(Number := 61,
                  Operation := 2,
                  Signal := #r,
                  Preset := #a1);
   // PB20, STEP 5 network 5
   #r := ((NOT "ROLL_IO".Input[7, 2]) AND "ROLL_State".S5Timers[55].Q);
   IF #r THEN
       "ROLL_State".M[8, 2] := TRUE;
   END_IF;
   #r := "ROLL_State".M[3, 1];
   IF #r THEN
       "ROLL_State".M[8, 2] := FALSE;
   END_IF;
   // PB20, STEP 5 network 6
   #a2 := #a1;
   #a1 := "ROLL_GetDW"(DbNumber := #activeDataBlock, Index := 55);
   #r := ((NOT "ROLL_IO".Input[7, 2]) AND (NOT "ROLL_State".M[8, 2]) AND "ROLL_State".M[4, 1]);
   "ROLL_TimerOp"(Number := 55,
                  Operation := 0,
                  Signal := #r,
                  Preset := #a1);
   // PB20, STEP 5 network 7
   #r := ((NOT "ROLL_IO".Input[7, 3]) AND "ROLL_IO".Output[21, 6] AND "ROLL_State".S5Timers[60].Q);
   IF #r THEN
       "ROLL_State".M[8, 3] := TRUE;
   END_IF;
   #r := "ROLL_State".M[3, 1];
   IF #r THEN
       "ROLL_State".M[8, 3] := FALSE;
   END_IF;
   // PB20, STEP 5 network 8
   #a2 := #a1;
   #a1 := "ROLL_GetDW"(DbNumber := #activeDataBlock, Index := 60);
   #r := ((NOT "ROLL_IO".Input[7, 3]) AND "ROLL_IO".Output[21, 6] AND "ROLL_IO".Input[3, 1]);
   "ROLL_TimerOp"(Number := 60,
                  Operation := 0,
                  Signal := #r,
                  Preset := #a1);
   // PB20, STEP 5 network 9
   #a2 := #a1;
   #a1 := W#16#2010;
   #r := (NOT "ROLL_IO".Input[7, 4]);
   "ROLL_TimerOp"(Number := 88,
                  Operation := 0,
                  Signal := #r,
                  Preset := #a1);
   // PB20, STEP 5 network 10
   #r := ((NOT "ROLL_IO".Input[7, 4]) AND "ROLL_State".M[4, 1] AND "ROLL_State".S5Timers[88].Q);
   "ROLL_State".M[8, 4] := #r;
   // PB20, STEP 5 network 11
   #r := (("ROLL_State".M[25, 0] OR "ROLL_State".M[25, 1]) AND "ROLL_IO".Input[0, 1] AND "ROLL_State".M[190, 6] AND "ROLL_State".M[4, 1] AND "ROLL_State".S5Timers[96].Q);
   IF #r THEN
       "ROLL_State".M[8, 5] := TRUE;
   END_IF;
   #r := "ROLL_State".M[3, 1];
   IF #r THEN
       "ROLL_State".M[8, 5] := FALSE;
   END_IF;
   // PB20, STEP 5 network 12
   #r := ((NOT "ROLL_IO".Input[9, 0]) AND ("ROLL_IO".Input[1, 6] OR "ROLL_IO".Input[1, 7]) AND "ROLL_IO".Input[9, 6]);
   IF #r THEN
       "ROLL_State".M[12, 4] := TRUE;
   END_IF;
   #r := "ROLL_State".M[3, 1];
   IF #r THEN
       "ROLL_State".M[12, 4] := FALSE;
   END_IF;
   // PB20, STEP 5 network 13
   #r := ((NOT "ROLL_IO".Input[9, 3]) AND ("ROLL_IO".Input[1, 6] OR "ROLL_IO".Input[1, 7]) AND "ROLL_IO".Input[9, 6]);
   IF #r THEN
       "ROLL_State".M[12, 5] := TRUE;
   END_IF;
   #r := "ROLL_State".M[3, 1];
   IF #r THEN
       "ROLL_State".M[12, 5] := FALSE;
   END_IF;
   // PB20, STEP 5 network 14
   #r := ((NOT "ROLL_IO".Input[9, 7]) AND ("ROLL_IO".Input[1, 6] OR "ROLL_IO".Input[1, 7]));
   IF #r THEN
       "ROLL_State".M[12, 6] := TRUE;
   END_IF;
   #r := "ROLL_State".M[3, 1];
   IF #r THEN
       "ROLL_State".M[12, 6] := FALSE;
   END_IF;
   // PB20, STEP 5 network 15
   #r := (NOT "ROLL_IO".Input[9, 6]);
   IF #r THEN
       "ROLL_State".M[12, 7] := TRUE;
   END_IF;
   #r := ("ROLL_IO".Input[9, 6] AND "ROLL_State".M[3, 1]);
   IF #r THEN
       "ROLL_State".M[12, 7] := FALSE;
   END_IF;
   // PB20, STEP 5 network 16
   #a2 := #a1;
   #a1 := "ROLL_GetDW"(DbNumber := #activeDataBlock, Index := 56);
   #r := (NOT "ROLL_IO".Input[7, 1]);
   "ROLL_TimerOp"(Number := 56,
                  Operation := 1,
                  Signal := #r,
                  Preset := #a1);
   // PB20, STEP 5 network 17
   #a2 := #a1;
   #a1 := "ROLL_GetDW"(DbNumber := #activeDataBlock, Index := 65);
   #r := (NOT "ROLL_IO".Input[7, 3]);
   "ROLL_TimerOp"(Number := 65,
                  Operation := 0,
                  Signal := #r,
                  Preset := #a1);
   // PB20, STEP 5 network 18
   #a2 := #a1;
   #a1 := W#16#2020;
   #r := "ROLL_IO".Input[7, 3];
   "ROLL_TimerOp"(Number := 66,
                  Operation := 1,
                  Signal := #r,
                  Preset := #a1);
   // PB20, STEP 5 network 19
   #a2 := #a1;
   #a1 := "ROLL_GetDW"(DbNumber := #activeDataBlock, Index := 67);
   #r := ("ROLL_IO".Input[7, 3] AND "ROLL_State".M[150, 1]);
   "ROLL_TimerOp"(Number := 67,
                  Operation := 0,
                  Signal := #r,
                  Preset := #a1);
   // PB20, STEP 5 network 20
   #a2 := #a1;
   #a1 := W#16#2005;
   #r := (NOT "ROLL_IO".Input[7, 5]);
   "ROLL_TimerOp"(Number := 96,
                  Operation := 0,
                  Signal := #r,
                  Preset := #a1);
   // PB20, STEP 5 network 21
   #a2 := #a1;
   #a1 := W#16#2030;
   #r := "ROLL_IO".Input[7, 5];
   "ROLL_TimerOp"(Number := 97,
                  Operation := 0,
                  Signal := #r,
                  Preset := #a1);
   // PB20, STEP 5 network 22
   #r := (((NOT "ROLL_IO".Output[18, 5]) AND "ROLL_IO".Output[18, 4]) OR ((NOT "ROLL_IO".Output[18, 7]) AND "ROLL_IO".Output[18, 6]));
   "ROLL_State".M[149, 6] := #r;
   // PB20, STEP 5 network 23
   #a2 := #a1;
   #a1 := W#16#1010;
   #r := "ROLL_State".M[148, 4];
   "ROLL_TimerOp"(Number := 89,
                  Operation := 0,
                  Signal := #r,
                  Preset := #a1);
   // PB20, STEP 5 network 24
   #r := "ROLL_State".M[149, 6];
   IF #r THEN
       "ROLL_State".M[148, 4] := TRUE;
   END_IF;
   #r := "ROLL_State".S5Timers[89].Q;
   IF #r THEN
       "ROLL_State".M[148, 4] := FALSE;
   END_IF;
   // PB20, STEP 5 network 25
   #r := ("ROLL_IO".Input[8, 0] AND "ROLL_State".S5Timers[70].Q);
   "ROLL_State".M[147, 0] := #r;
   // PB20, STEP 5 network 26
   #a2 := #a1;
   #a1 := "ROLL_GetDW"(DbNumber := #activeDataBlock, Index := 75);
   #r := (NOT "ROLL_State".M[147, 0]);
   "ROLL_TimerOp"(Number := 75,
                  Operation := 0,
                  Signal := #r,
                  Preset := #a1);
   // PB20, STEP 5 network 27
   #r := "ROLL_State".M[0, 3];
   "ROLL_State".M[147, 1] := #r;
   // PB20, STEP 5 network 28
   #r := ("ROLL_IO".Input[8, 2] AND "ROLL_State".S5Timers[72].Q);
   "ROLL_State".M[147, 2] := #r;
   // PB20, STEP 5 network 29
   #a2 := #a1;
   #a1 := "ROLL_GetDW"(DbNumber := #activeDataBlock, Index := 77);
   #r := (NOT "ROLL_State".M[147, 2]);
   "ROLL_TimerOp"(Number := 77,
                  Operation := 0,
                  Signal := #r,
                  Preset := #a1);
   // PB20, STEP 5 network 30
   #r := "ROLL_State".M[0, 3];
   "ROLL_State".M[149, 0] := #r;
   // PB20, STEP 5 network 31
   #r := ("ROLL_State".M[147, 0] OR "ROLL_State".M[147, 2]);
   "ROLL_State".M[149, 1] := #r;
   // PB20, STEP 5 network 32
   #r := "ROLL_State".M[0, 3];
   "ROLL_State".M[149, 2] := #r;
   // PB20, STEP 5 network 33
   #r := ("ROLL_State".M[147, 0] AND "ROLL_State".M[147, 2]);
   "ROLL_State".M[149, 3] := #r;
   // PB20, STEP 5 network 34
   #r := ((NOT "ROLL_State".M[12, 6]) AND (NOT "ROLL_State".M[12, 7]) AND (NOT "ROLL_State".M[13, 4]) AND (NOT "ROLL_State".M[6, 0]) AND (NOT "ROLL_State".M[6, 2]) AND (NOT "ROLL_State".M[8, 2]) AND ("ROLL_IO".Input[1, 6] OR "ROLL_IO".Input[1, 7]) AND "ROLL_IO".Input[3, 1] AND "ROLL_IO".Input[7, 4] AND "ROLL_IO".Input[9, 6] AND "ROLL_IO".Input[9, 7] AND "ROLL_State".S5Timers[66].Q);
   "ROLL_State".M[150, 2] := #r;
   // PB20, STEP 5 network 35
   #r := ((NOT "ROLL_IO".Input[9, 2]) AND (NOT "ROLL_State".M[12, 4]) AND ("ROLL_IO".Output[18, 4] OR "ROLL_IO".Input[9, 1]) AND ("ROLL_State".M[149, 0] OR "ROLL_State".M[149, 1] OR "ROLL_State".M[149, 2] OR "ROLL_State".M[149, 3]) AND "ROLL_IO".Input[9, 0] AND "ROLL_State".M[150, 2]);
   "ROLL_IO".Output[18, 4] := #r;
   // PB20, STEP 5 network 36
   #r := ((NOT "ROLL_IO".Input[9, 2]) AND (NOT "ROLL_State".M[12, 4]) AND ("ROLL_IO".Output[18, 4] OR "ROLL_IO".Output[18, 5] OR "ROLL_IO".Input[9, 1]) AND ("ROLL_State".M[149, 2] OR "ROLL_State".M[149, 3]) AND "ROLL_IO".Input[9, 0] AND "ROLL_State".M[150, 2]);
   "ROLL_IO".Output[18, 5] := #r;
   // PB20, STEP 5 network 37
   #r := ((NOT "ROLL_IO".Input[9, 5]) AND (NOT "ROLL_State".M[12, 5]) AND ("ROLL_IO".Output[18, 6] OR "ROLL_IO".Input[9, 4]) AND ("ROLL_State".M[149, 1] OR "ROLL_State".M[149, 2] OR "ROLL_State".M[149, 3]) AND "ROLL_IO".Input[9, 3] AND "ROLL_State".M[150, 2]);
   "ROLL_IO".Output[18, 6] := #r;
   // PB20, STEP 5 network 38
   #r := ((NOT "ROLL_IO".Input[9, 5]) AND (NOT "ROLL_State".M[12, 5]) AND ("ROLL_IO".Output[18, 6] OR "ROLL_IO".Output[18, 7] OR "ROLL_IO".Input[9, 4]) AND "ROLL_IO".Input[9, 3] AND "ROLL_State".M[149, 3] AND "ROLL_State".M[150, 2]);
   "ROLL_IO".Output[18, 7] := #r;
   // PB20, STEP 5 network 39
   #r := ((NOT "ROLL_State".M[147, 0]) AND "ROLL_State".M[147, 2] AND "ROLL_State".S5Timers[75].Q);
   "ROLL_IO".Output[21, 0] := #r;
   // PB20, STEP 5 network 40
   #r := ((NOT "ROLL_State".M[147, 2]) AND "ROLL_State".M[147, 0] AND "ROLL_State".S5Timers[77].Q);
   "ROLL_IO".Output[21, 2] := #r;
   // PB20, STEP 5 network 41
   #r := "ROLL_State".M[190, 6];
   IF #r THEN
       "ROLL_State".M[150, 0] := TRUE;
   END_IF;
   #r := ((NOT "ROLL_IO".Input[0, 1]) OR (NOT "ROLL_IO".Input[7, 1]) OR (NOT "ROLL_IO".Input[7, 2]) OR (NOT "ROLL_State".M[27, 5]) OR "ROLL_IO".Input[7, 3] OR "ROLL_State".M[190, 5]);
   IF #r THEN
       "ROLL_State".M[150, 0] := FALSE;
   END_IF;
   // PB20, STEP 5 network 42
   #a2 := #a1;
   #a1 := W#16#2020;
   #r := "ROLL_IO".Input[7, 1];
   "ROLL_TimerOp"(Number := 57,
                  Operation := 1,
                  Signal := #r,
                  Preset := #a1);
   // PB20, STEP 5 network 43
   #r := ((NOT "ROLL_State".M[13, 4]) AND (NOT "ROLL_State".S5Timers[61].Q) AND (((NOT "ROLL_IO".Input[7, 3]) AND "ROLL_State".S5Timers[65].Q) OR ((NOT "ROLL_State".S5Timers[67].Q) AND "ROLL_State".M[150, 1])) AND "ROLL_IO".Input[0, 2] AND "ROLL_IO".Input[3, 1] AND "ROLL_IO".Input[7, 2] AND "ROLL_State".S5Timers[57].Q);
   "ROLL_State".M[150, 1] := #r;
   // PB20, STEP 5 network 44
   #r := ("ROLL_State".M[150, 0] OR "ROLL_State".M[150, 1]);
   "ROLL_IO".Output[21, 6] := #r;
   // PB20, STEP 5 network 45
   #r := ((((NOT "ROLL_IO".Input[7, 4]) AND "ROLL_IO".Input[7, 5]) OR ((NOT "ROLL_State".S5Timers[106].Q) AND "ROLL_State".M[148, 6]) OR (NOT "ROLL_IO".Input[7, 1])) AND "ROLL_IO".Input[0, 2] AND "ROLL_IO".Input[1, 6] AND "ROLL_IO".Input[7, 0]);
   "ROLL_State".M[148, 6] := #r;
   // PB20, STEP 5 network 46
   #r := (((NOT "ROLL_State".M[151, 0]) AND (NOT "ROLL_State".M[151, 1]) AND (NOT "ROLL_State".M[151, 2]) AND (NOT "ROLL_State".M[151, 3])) OR ((NOT "ROLL_State".M[152, 3]) AND "ROLL_State".M[151, 3] AND "ROLL_State".M[153, 3] AND "ROLL_State".S5Timers[105].Q));
   IF #r THEN
       "ROLL_State".M[151, 0] := TRUE;
   END_IF;
   #r := ("ROLL_State".M[151, 1] OR "ROLL_State".M[151, 2]);
   IF #r THEN
       "ROLL_State".M[151, 0] := FALSE;
   END_IF;
   // PB20, STEP 5 network 47
   #a2 := #a1;
   #a1 := "ROLL_GetDW"(DbNumber := #activeDataBlock, Index := 102);
   #r := "ROLL_State".M[151, 0];
   "ROLL_TimerOp"(Number := 102,
                  Operation := 0,
                  Signal := #r,
                  Preset := #a1);
   // PB20, STEP 5 network 48
   #r := ((NOT "ROLL_State".S5Timers[106].Q) AND "ROLL_State".M[151, 0]);
   IF #r THEN
       "ROLL_State".M[152, 0] := TRUE;
   END_IF;
   #r := ((NOT "ROLL_State".M[148, 6]) OR "ROLL_State".S5Timers[106].Q);
   IF #r THEN
       "ROLL_State".M[152, 0] := FALSE;
   END_IF;
   // PB20, STEP 5 network 49
   #r := ("ROLL_IO".Output[21, 5] AND "ROLL_State".M[152, 0]);
   IF #r THEN
       "ROLL_State".M[153, 0] := TRUE;
   END_IF;
   #r := (NOT "ROLL_State".M[151, 0]);
   IF #r THEN
       "ROLL_State".M[153, 0] := FALSE;
   END_IF;
   // PB20, STEP 5 network 50
   #r := ((NOT "ROLL_State".M[152, 0]) AND "ROLL_State".M[151, 0] AND "ROLL_State".M[153, 0] AND "ROLL_State".S5Timers[102].Q);
   IF #r THEN
       "ROLL_State".M[151, 1] := TRUE;
   END_IF;
   #r := "ROLL_State".M[151, 2];
   IF #r THEN
       "ROLL_State".M[151, 1] := FALSE;
   END_IF;
   // PB20, STEP 5 network 51
   #a2 := #a1;
   #a1 := "ROLL_GetDW"(DbNumber := #activeDataBlock, Index := 103);
   #r := "ROLL_State".M[151, 1];
   "ROLL_TimerOp"(Number := 103,
                  Operation := 0,
                  Signal := #r,
                  Preset := #a1);
   // PB20, STEP 5 network 52
   #r := ((NOT "ROLL_State".S5Timers[106].Q) AND "ROLL_State".M[151, 1]);
   IF #r THEN
       "ROLL_State".M[152, 1] := TRUE;
   END_IF;
   #r := ((NOT "ROLL_State".M[148, 6]) OR "ROLL_State".S5Timers[106].Q);
   IF #r THEN
       "ROLL_State".M[152, 1] := FALSE;
   END_IF;
   // PB20, STEP 5 network 53
   #r := ("ROLL_IO".Output[20, 6] AND "ROLL_State".M[152, 1]);
   IF #r THEN
       "ROLL_State".M[153, 1] := TRUE;
   END_IF;
   #r := (NOT "ROLL_State".M[151, 1]);
   IF #r THEN
       "ROLL_State".M[153, 1] := FALSE;
   END_IF;
   // PB20, STEP 5 network 54
   #r := ((NOT "ROLL_State".M[152, 1]) AND "ROLL_State".M[151, 1] AND "ROLL_State".M[153, 1] AND "ROLL_State".S5Timers[103].Q);
   IF #r THEN
       "ROLL_State".M[151, 2] := TRUE;
   END_IF;
   #r := "ROLL_State".M[151, 3];
   IF #r THEN
       "ROLL_State".M[151, 2] := FALSE;
   END_IF;
   // PB20, STEP 5 network 55
   #a2 := #a1;
   #a1 := W#16#0002;
   #r := "ROLL_State".M[151, 2];
   "ROLL_TimerOp"(Number := 104,
                  Operation := 0,
                  Signal := #r,
                  Preset := #a1);
   // PB20, STEP 5 network 56
   #r := ((NOT "ROLL_State".S5Timers[106].Q) AND "ROLL_State".M[151, 2]);
   IF #r THEN
       "ROLL_State".M[152, 2] := TRUE;
   END_IF;
   #r := ((NOT "ROLL_State".M[148, 6]) OR "ROLL_State".S5Timers[106].Q);
   IF #r THEN
       "ROLL_State".M[152, 2] := FALSE;
   END_IF;
   // PB20, STEP 5 network 57
   #r := ("ROLL_State".M[0, 4] AND "ROLL_State".M[152, 2]);
   IF #r THEN
       "ROLL_State".M[153, 2] := TRUE;
   END_IF;
   #r := (NOT "ROLL_State".M[151, 2]);
   IF #r THEN
       "ROLL_State".M[153, 2] := FALSE;
   END_IF;
   // PB20, STEP 5 network 58
   #r := ((NOT "ROLL_State".M[152, 2]) AND "ROLL_State".M[151, 2] AND "ROLL_State".M[153, 2] AND "ROLL_State".S5Timers[104].Q);
   IF #r THEN
       "ROLL_State".M[151, 3] := TRUE;
   END_IF;
   #r := "ROLL_State".M[151, 0];
   IF #r THEN
       "ROLL_State".M[151, 3] := FALSE;
   END_IF;
   // PB20, STEP 5 network 59
   #a2 := #a1;
   #a1 := W#16#0002;
   #r := "ROLL_State".M[151, 3];
   "ROLL_TimerOp"(Number := 105,
                  Operation := 0,
                  Signal := #r,
                  Preset := #a1);
   // PB20, STEP 5 network 60
   #r := ((NOT "ROLL_State".S5Timers[106].Q) AND "ROLL_State".M[151, 3]);
   IF #r THEN
       "ROLL_State".M[152, 3] := TRUE;
   END_IF;
   #r := ((NOT "ROLL_State".M[148, 6]) OR "ROLL_State".S5Timers[106].Q);
   IF #r THEN
       "ROLL_State".M[152, 3] := FALSE;
   END_IF;
   // PB20, STEP 5 network 61
   #r := ("ROLL_State".M[0, 4] AND "ROLL_State".M[152, 3]);
   IF #r THEN
       "ROLL_State".M[153, 3] := TRUE;
   END_IF;
   #r := (NOT "ROLL_State".M[151, 3]);
   IF #r THEN
       "ROLL_State".M[153, 3] := FALSE;
   END_IF;
   // PB20, STEP 5 network 62
   #a2 := #a1;
   #a1 := W#16#2010;
   #r := ("ROLL_State".M[152, 0] OR "ROLL_State".M[152, 1] OR "ROLL_State".M[152, 2] OR "ROLL_State".M[152, 3]);
   "ROLL_TimerOp"(Number := 106,
                  Operation := 0,
                  Signal := #r,
                  Preset := #a1);
   // PB20, STEP 5 network 63
   #r := ((NOT "ROLL_IO".Output[21, 4]) AND "ROLL_IO".Output[19, 5] AND "ROLL_State".M[152, 0]);
   "ROLL_IO".Output[21, 5] := #r;
   // PB20, STEP 5 network 64
   #r := "ROLL_State".M[152, 1];
   "ROLL_State".M[240, 0] := #r;
   // PB20, STEP 5 network 65
   #r := ((NOT "ROLL_IO".Output[21, 5]) AND "ROLL_State".M[152, 2]);
   "ROLL_State".M[240, 0] := #r;
   // PB20, STEP 5 network 66
   #r := "ROLL_State".M[152, 3];
   "ROLL_State".M[240, 0] := #r;
   // PB20, STEP 5 network 67
   #a2 := #a1;
   #a1 := "ROLL_GetDW"(DbNumber := #activeDataBlock, Index := 107);
   #r := ("ROLL_IO".Output[21, 6] AND "ROLL_IO".Input[0, 2]);
   "ROLL_TimerOp"(Number := 107,
                  Operation := 1,
                  Signal := #r,
                  Preset := #a1);
   // PB20, STEP 5 network 68
   #r := ((("ROLL_IO".Output[21, 6] OR "ROLL_State".S5Timers[107].Q) AND "ROLL_IO".Input[0, 2]) OR ("ROLL_IO".Input[0, 1] AND "ROLL_State".M[190, 6] AND "ROLL_State".M[26, 6]));
   "ROLL_IO".Output[20, 5] := #r;
   // PB20, STEP 5 network 69
   RETURN;
END_FUNCTION

FUNCTION "ROLL_PB21" : Void   // FC29, SCL
{ S7_Optimized_Access := 'TRUE' }
VERSION : 0.1
// stored: AutoNumber true, IsIECCheckEnabled false, SetENOAutomatically false, UDAEnableTagReadback false
   VAR_TEMP
      r : Bool;
      a1 : Word;
      a2 : Word;
      activeDataBlock : Int;
      comparisonResults : Array[0..0] of Bool;
   END_VAR
BEGIN

   #r := FALSE;
   #a1 := W#16#0000;
   #a2 := W#16#0000;
   #activeDataBlock := 0;
   // PB21, STEP 5 network 1
   #activeDataBlock := 15;
   // PB21, STEP 5 network 2
   #r := ((NOT "ROLL_IO".Input[3, 6]) AND (NOT "ROLL_State".M[13, 1]) AND (NOT "ROLL_State".M[5, 6]));
   "ROLL_State".M[99, 7] := #r;
   // PB21, STEP 5 network 3
   #r := ((NOT "ROLL_State".M[13, 3]) AND (NOT "ROLL_State".M[16, 6]) AND (NOT "ROLL_State".M[6, 0]) AND (NOT "ROLL_State".M[6, 2]) AND "ROLL_IO".Input[3, 0] AND "ROLL_IO".Input[5, 0] AND "ROLL_IO".Input[5, 2] AND "ROLL_IO".Input[5, 4]);
   "ROLL_State".M[100, 0] := #r;
   // PB21, STEP 5 network 4
   #r := "ROLL_State".M[190, 6];
   IF #r THEN
       "ROLL_State".M[100, 1] := TRUE;
   END_IF;
   #r := (((NOT "ROLL_State".M[190, 6]) AND "ROLL_IO".Input[5, 3]) OR (NOT "ROLL_IO".Input[0, 1]) OR (NOT "ROLL_State".M[0, 3]) OR (NOT "ROLL_State".M[100, 0]) OR "ROLL_State".M[190, 5]);
   IF #r THEN
       "ROLL_State".M[100, 1] := FALSE;
   END_IF;
   // PB21, STEP 5 network 5
   #r := "ROLL_State".M[190, 6];
   IF #r THEN
       "ROLL_State".M[100, 2] := TRUE;
   END_IF;
   #r := (("ROLL_IO".Input[5, 3] AND "ROLL_IO".Input[5, 6]) OR (NOT "ROLL_IO".Input[0, 1]) OR (NOT "ROLL_State".M[0, 3]) OR (NOT "ROLL_State".M[100, 0]) OR "ROLL_State".M[190, 5]);
   IF #r THEN
       "ROLL_State".M[100, 2] := FALSE;
   END_IF;
   // PB21, STEP 5 network 6
   #r := "ROLL_State".M[190, 6];
   IF #r THEN
       "ROLL_State".M[100, 3] := TRUE;
   END_IF;
   #r := (((NOT "ROLL_IO".Input[7, 5]) AND (NOT "ROLL_State".M[190, 6])) OR (NOT "ROLL_IO".Input[0, 1]) OR (NOT "ROLL_State".M[0, 3]) OR (NOT "ROLL_State".M[100, 0]) OR "ROLL_State".M[190, 5] OR "ROLL_State".M[5, 6] OR "ROLL_State".M[8, 5]);
   IF #r THEN
       "ROLL_State".M[100, 3] := FALSE;
   END_IF;
   // PB21, STEP 5 network 7
   #r := "ROLL_State".M[190, 6];
   IF #r THEN
       "ROLL_State".M[100, 4] := TRUE;
   END_IF;
   #r := (((NOT "ROLL_State".M[100, 0]) AND (NOT "ROLL_State".M[190, 6])) OR (NOT "ROLL_IO".Input[0, 1]) OR (NOT "ROLL_State".M[0, 3]) OR (NOT "ROLL_State".M[99, 7]) OR "ROLL_State".M[190, 5]);
   IF #r THEN
       "ROLL_State".M[100, 4] := FALSE;
   END_IF;
   // PB21, STEP 5 network 8
   #r := ((NOT "ROLL_State".M[31, 5]) AND (NOT "ROLL_State".M[5, 6]) AND ((NOT "ROLL_IO".Input[5, 6]) OR (NOT "ROLL_State".S5Timers[70].Q)) AND "ROLL_IO".Input[0, 2] AND "ROLL_IO".Input[3, 1] AND "ROLL_State".M[100, 0]);
   "ROLL_State".M[100, 5] := #r;
   // PB21, STEP 5 network 9
   #r := ((("ROLL_IO".Input[7, 5] AND "ROLL_State".S5Timers[97].Q) OR (NOT "ROLL_State".S5Timers[96].Q)) AND "ROLL_State".M[0, 3] AND "ROLL_State".M[100, 5]);
   "ROLL_State".M[100, 6] := #r;
   // PB21, STEP 5 network 10
   #r := ((((NOT "ROLL_IO".Input[7, 5]) AND "ROLL_State".S5Timers[96].Q) OR (NOT "ROLL_State".S5Timers[97].Q)) AND "ROLL_State".M[0, 3] AND "ROLL_State".M[100, 5]);
   "ROLL_State".M[100, 7] := #r;
   // PB21, STEP 5 network 11
   #r := "ROLL_State".M[190, 6];
   IF #r THEN
       "ROLL_State".M[101, 1] := TRUE;
   END_IF;
   #r := (((NOT "ROLL_State".M[190, 6]) AND "ROLL_IO".Input[5, 3] AND "ROLL_IO".Input[5, 6] AND "ROLL_IO".Input[6, 0]) OR (NOT "ROLL_IO".Input[0, 1]) OR (NOT "ROLL_State".M[0, 3]) OR (NOT "ROLL_State".M[100, 0]) OR "ROLL_State".M[190, 5]);
   IF #r THEN
       "ROLL_State".M[101, 1] := FALSE;
   END_IF;
   // PB21, STEP 5 network 12
   #r := "ROLL_State".M[190, 6];
   IF #r THEN
       "ROLL_State".M[101, 2] := TRUE;
   END_IF;
   #r := (((NOT "ROLL_State".M[190, 6]) AND "ROLL_IO".Input[5, 3] AND "ROLL_IO".Input[5, 6] AND "ROLL_IO".Input[6, 0]) OR (NOT "ROLL_IO".Input[0, 1]) OR (NOT "ROLL_State".M[0, 3]) OR (NOT "ROLL_State".M[100, 0]) OR "ROLL_State".M[190, 5]);
   IF #r THEN
       "ROLL_State".M[101, 2] := FALSE;
   END_IF;
   // PB21, STEP 5 network 13
   #r := "ROLL_State".M[190, 6];
   IF #r THEN
       "ROLL_State".M[101, 3] := TRUE;
   END_IF;
   #r := (((NOT "ROLL_State".M[190, 6]) AND ((NOT "ROLL_IO".Input[7, 5]) OR "ROLL_IO".Input[6, 0])) OR (NOT "ROLL_IO".Input[0, 1]) OR (NOT "ROLL_State".M[0, 3]) OR (NOT "ROLL_State".M[100, 0]) OR "ROLL_State".M[190, 5] OR "ROLL_State".M[5, 6] OR "ROLL_State".M[8, 5]);
   IF #r THEN
       "ROLL_State".M[101, 3] := FALSE;
   END_IF;
   // PB21, STEP 5 network 14
   #r := "ROLL_State".M[190, 6];
   IF #r THEN
       "ROLL_State".M[101, 4] := TRUE;
   END_IF;
   #r := (((NOT "ROLL_State".M[190, 6]) AND "ROLL_IO".Input[6, 0]) OR (NOT "ROLL_IO".Input[0, 1]) OR (NOT "ROLL_State".M[0, 3]) OR (NOT "ROLL_State".M[100, 0]) OR (NOT "ROLL_State".M[99, 7]) OR "ROLL_State".M[190, 5]);
   IF #r THEN
       "ROLL_State".M[101, 4] := FALSE;
   END_IF;
   // PB21, STEP 5 network 15
   #a2 := #a1;
   #a1 := W#16#2005;
   #r := "ROLL_IO".Input[6, 0];
   "ROLL_TimerOp"(Number := 121,
                  Operation := 0,
                  Signal := #r,
                  Preset := #a1);
   // PB21, STEP 5 network 16
   #r := ((NOT "ROLL_State".M[31, 5]) AND (NOT "ROLL_State".M[5, 6]) AND (((NOT "ROLL_State".S5Timers[121].Q) AND "ROLL_State".M[101, 5]) OR (NOT "ROLL_IO".Input[6, 0])) AND "ROLL_IO".Input[0, 2] AND "ROLL_IO".Input[3, 1] AND "ROLL_State".M[100, 0]);
   "ROLL_State".M[101, 5] := #r;
   // PB21, STEP 5 network 17
   #r := ((("ROLL_IO".Input[7, 5] AND "ROLL_State".S5Timers[97].Q) OR (NOT "ROLL_State".S5Timers[96].Q)) AND "ROLL_State".M[101, 5]);
   "ROLL_State".M[101, 6] := #r;
   // PB21, STEP 5 network 18
   #r := ((((NOT "ROLL_IO".Input[7, 5]) AND "ROLL_State".S5Timers[96].Q) OR (NOT "ROLL_State".S5Timers[97].Q)) AND "ROLL_State".M[101, 5]);
   "ROLL_State".M[101, 7] := #r;
   // PB21, STEP 5 network 19
   #r := "ROLL_State".M[190, 6];
   IF #r THEN
       "ROLL_State".M[102, 1] := TRUE;
   END_IF;
   #r := (((NOT "ROLL_State".M[190, 6]) AND "ROLL_IO".Input[5, 3] AND "ROLL_IO".Input[5, 6] AND "ROLL_IO".Input[6, 0] AND "ROLL_IO".Input[6, 2]) OR (NOT "ROLL_IO".Input[0, 1]) OR (NOT "ROLL_State".M[0, 3]) OR (NOT "ROLL_State".M[100, 0]) OR "ROLL_State".M[190, 5]);
   IF #r THEN
       "ROLL_State".M[102, 1] := FALSE;
   END_IF;
   // PB21, STEP 5 network 20
   #r := "ROLL_State".M[190, 6];
   IF #r THEN
       "ROLL_State".M[102, 2] := TRUE;
   END_IF;
   #r := (((NOT "ROLL_State".M[190, 6]) AND "ROLL_IO".Input[6, 2]) OR (NOT "ROLL_IO".Input[0, 1]) OR (NOT "ROLL_State".M[0, 3]) OR (NOT "ROLL_State".M[100, 0]) OR "ROLL_State".M[190, 5]);
   IF #r THEN
       "ROLL_State".M[102, 2] := FALSE;
   END_IF;
   // PB21, STEP 5 network 21
   #r := "ROLL_State".M[190, 6];
   IF #r THEN
       "ROLL_State".M[102, 3] := TRUE;
   END_IF;
   #r := (((NOT "ROLL_State".M[190, 6]) AND ((NOT "ROLL_IO".Input[7, 5]) OR "ROLL_IO".Input[6, 2])) OR (NOT "ROLL_IO".Input[0, 1]) OR (NOT "ROLL_State".M[0, 3]) OR (NOT "ROLL_State".M[100, 0]) OR "ROLL_State".M[190, 5] OR "ROLL_State".M[5, 6] OR "ROLL_State".M[8, 5]);
   IF #r THEN
       "ROLL_State".M[102, 3] := FALSE;
   END_IF;
   // PB21, STEP 5 network 22
   #r := "ROLL_State".M[190, 6];
   IF #r THEN
       "ROLL_State".M[102, 4] := TRUE;
   END_IF;
   #r := (((NOT "ROLL_State".M[190, 6]) AND "ROLL_IO".Input[6, 2]) OR (NOT "ROLL_IO".Input[0, 1]) OR (NOT "ROLL_State".M[0, 3]) OR (NOT "ROLL_State".M[100, 0]) OR (NOT "ROLL_State".M[99, 7]) OR "ROLL_State".M[190, 5]);
   IF #r THEN
       "ROLL_State".M[102, 4] := FALSE;
   END_IF;
   // PB21, STEP 5 network 23
   #r := ((NOT "ROLL_State".M[31, 5]) AND (NOT "ROLL_State".M[5, 6]) AND (NOT "ROLL_State".S5Timers[72].Q) AND "ROLL_IO".Input[0, 2] AND "ROLL_IO".Input[3, 1] AND "ROLL_State".M[100, 0]);
   "ROLL_State".M[102, 5] := #r;
   // PB21, STEP 5 network 24
   #r := ((("ROLL_IO".Input[7, 5] AND "ROLL_State".S5Timers[97].Q) OR (NOT "ROLL_State".S5Timers[96].Q)) AND "ROLL_State".M[0, 3] AND "ROLL_State".M[102, 5]);
   "ROLL_State".M[102, 6] := #r;
   // PB21, STEP 5 network 25
   #r := ((((NOT "ROLL_IO".Input[7, 5]) AND "ROLL_State".S5Timers[96].Q) OR (NOT "ROLL_State".S5Timers[97].Q) OR "ROLL_State".M[0, 4]) AND "ROLL_State".M[102, 5]);
   "ROLL_State".M[102, 7] := #r;
   // PB21, STEP 5 network 26
   #r := "ROLL_State".M[190, 6];
   IF #r THEN
       "ROLL_State".M[105, 1] := TRUE;
   END_IF;
   #r := (((NOT "ROLL_State".M[190, 6]) AND "ROLL_State".M[0, 4]) OR (NOT "ROLL_IO".Input[0, 1]) OR (NOT "ROLL_State".M[0, 3]) OR (NOT "ROLL_State".M[100, 0]) OR "ROLL_State".M[190, 5]);
   IF #r THEN
       "ROLL_State".M[105, 1] := FALSE;
   END_IF;
   // PB21, STEP 5 network 27
   #r := "ROLL_State".M[190, 6];
   IF #r THEN
       "ROLL_State".M[105, 2] := TRUE;
   END_IF;
   #r := ((NOT "ROLL_IO".Input[0, 1]) OR (NOT "ROLL_State".M[0, 3]) OR (NOT "ROLL_State".M[100, 0]) OR "ROLL_IO".Input[6, 2] OR "ROLL_State".M[190, 5]);
   IF #r THEN
       "ROLL_State".M[105, 2] := FALSE;
   END_IF;
   // PB21, STEP 5 network 28
   #r := "ROLL_State".M[190, 6];
   IF #r THEN
       "ROLL_State".M[105, 3] := TRUE;
   END_IF;
   #r := (((NOT "ROLL_State".M[190, 6]) AND ((NOT "ROLL_IO".Input[7, 5]) OR "ROLL_State".M[0, 4])) OR (NOT "ROLL_IO".Input[0, 1]) OR (NOT "ROLL_State".M[0, 3]) OR (NOT "ROLL_State".M[100, 0]) OR "ROLL_State".M[190, 5] OR "ROLL_State".M[5, 6] OR "ROLL_State".M[8, 5]);
   IF #r THEN
       "ROLL_State".M[105, 3] := FALSE;
   END_IF;
   // PB21, STEP 5 network 29
   #r := "ROLL_State".M[190, 6];
   IF #r THEN
       "ROLL_State".M[105, 4] := TRUE;
   END_IF;
   #r := (((NOT "ROLL_State".M[190, 6]) AND "ROLL_State".M[0, 4]) OR (NOT "ROLL_IO".Input[0, 1]) OR (NOT "ROLL_State".M[0, 3]) OR (NOT "ROLL_State".M[100, 0]) OR (NOT "ROLL_State".M[99, 7]) OR "ROLL_State".M[190, 5]);
   IF #r THEN
       "ROLL_State".M[105, 4] := FALSE;
   END_IF;
   // PB21, STEP 5 network 30
   #a2 := #a1;
   #a1 := W#16#2005;
   #r := "ROLL_State".M[0, 4];
   "ROLL_TimerOp"(Number := 120,
                  Operation := 0,
                  Signal := #r,
                  Preset := #a1);
   // PB21, STEP 5 network 31
   #r := ((NOT "ROLL_State".M[31, 5]) AND (NOT "ROLL_State".M[5, 6]) AND (((NOT "ROLL_State".S5Timers[120].Q) AND "ROLL_State".M[105, 5]) OR (NOT "ROLL_State".M[0, 4])) AND "ROLL_IO".Input[0, 2] AND "ROLL_IO".Input[3, 1] AND "ROLL_State".M[100, 0]);
   "ROLL_State".M[105, 5] := #r;
   // PB21, STEP 5 network 32
   #r := ((("ROLL_IO".Input[7, 5] AND "ROLL_State".S5Timers[97].Q) OR (NOT "ROLL_State".S5Timers[96].Q)) AND "ROLL_State".M[105, 5]);
   "ROLL_State".M[105, 6] := #r;
   // PB21, STEP 5 network 33
   #r := ((((NOT "ROLL_IO".Input[7, 5]) AND "ROLL_State".S5Timers[96].Q) OR (NOT "ROLL_State".S5Timers[97].Q)) AND "ROLL_State".M[105, 5]);
   "ROLL_State".M[105, 7] := #r;
   // PB21, STEP 5 network 34
   #r := ((((NOT "ROLL_IO".Input[5, 5]) AND ("ROLL_State".M[40, 5] OR "ROLL_State".M[42, 1]) AND "ROLL_State".M[31, 5]) OR (NOT "ROLL_IO".Input[5, 6])) AND "ROLL_IO".Input[0, 2] AND "ROLL_IO".Input[3, 1] AND "ROLL_State".M[100, 0]);
   "ROLL_State".M[103, 0] := #r;
   // PB21, STEP 5 network 35
   #r := (((NOT "ROLL_IO".Input[5, 3]) OR (NOT "ROLL_IO".Input[6, 0]) OR (NOT "ROLL_State".S5Timers[121].Q)) AND "ROLL_IO".Input[3, 1] AND "ROLL_State".M[100, 0] AND "ROLL_State".M[31, 5]);
   "ROLL_State".M[103, 3] := #r;
   // PB21, STEP 5 network 36
   #r := (((NOT "ROLL_IO".Input[5, 6]) AND "ROLL_IO".Input[0, 2]) OR (("ROLL_State".M[103, 0] OR "ROLL_State".M[103, 3]) AND "ROLL_State".S5Timers[62].Q AND "ROLL_State".S5Timers[97].Q));
   "ROLL_State".M[103, 1] := #r;
   // PB21, STEP 5 network 37
   #r := ((NOT "ROLL_IO".Input[6, 2]) AND "ROLL_IO".Input[3, 1] AND "ROLL_State".M[100, 0] AND "ROLL_State".M[31, 5]);
   "ROLL_State".M[103, 4] := #r;
   // PB21, STEP 5 network 38
   #a2 := #a1;
   #a1 := W#16#1050;
   #r := ("ROLL_IO".Output[22, 3] AND "ROLL_State".M[103, 4]);
   "ROLL_TimerOp"(Number := 119,
                  Operation := 1,
                  Signal := #r,
                  Preset := #a1);
   // PB21, STEP 5 network 39
   #r := (((("ROLL_State".M[103, 0] OR "ROLL_State".M[103, 3]) AND "ROLL_State".S5Timers[96].Q) OR "ROLL_State".M[103, 4] OR "ROLL_State".S5Timers[119].Q) AND "ROLL_State".S5Timers[62].Q);
   "ROLL_State".M[103, 2] := #r;
   // PB21, STEP 5 network 40
   #r := "ROLL_State".M[190, 6];
   IF #r THEN
       "ROLL_State".M[104, 0] := TRUE;
   END_IF;
   #r := (((NOT "ROLL_State".M[190, 6]) AND ((NOT "ROLL_IO".Input[5, 0]) OR (NOT "ROLL_IO".Input[5, 2]) OR (NOT "ROLL_IO".Input[5, 4]))) OR (NOT "ROLL_IO".Input[0, 1]) OR (NOT "ROLL_IO".Input[7, 0]) OR (NOT "ROLL_State".M[26, 5]) OR (NOT "ROLL_State".M[99, 7]) OR "ROLL_State".M[16, 6] OR "ROLL_State".M[190, 5]);
   IF #r THEN
       "ROLL_State".M[104, 0] := FALSE;
   END_IF;
   // PB21, STEP 5 network 41
   #r := "ROLL_State".M[190, 6];
   IF #r THEN
       "ROLL_State".M[104, 1] := TRUE;
   END_IF;
   #r := (((NOT "ROLL_State".M[190, 6]) AND ((NOT "ROLL_IO".Input[5, 0]) OR (NOT "ROLL_IO".Input[5, 2]) OR (NOT "ROLL_IO".Input[5, 4]))) OR (NOT "ROLL_IO".Input[0, 1]) OR (NOT "ROLL_State".M[26, 0]) OR (NOT "ROLL_State".M[99, 7]) OR "ROLL_State".M[16, 6] OR "ROLL_State".M[190, 5]);
   IF #r THEN
       "ROLL_State".M[104, 1] := FALSE;
   END_IF;
   // PB21, STEP 5 network 42
   #r := "ROLL_State".M[190, 6];
   IF #r THEN
       "ROLL_State".M[104, 4] := TRUE;
   END_IF;
   #r := (((NOT "ROLL_State".M[190, 6]) AND ((NOT "ROLL_IO".Input[5, 0]) OR (NOT "ROLL_IO".Input[5, 2]) OR (NOT "ROLL_IO".Input[5, 4]))) OR (NOT "ROLL_IO".Input[0, 1]) OR (NOT "ROLL_IO".Input[4, 7]) OR (NOT "ROLL_State".M[27, 4]) OR (NOT "ROLL_State".M[99, 7]) OR "ROLL_State".M[16, 6] OR "ROLL_State".M[190, 5]);
   IF #r THEN
       "ROLL_State".M[104, 4] := FALSE;
   END_IF;
   // PB21, STEP 5 network 43
   #r := "ROLL_State".M[190, 6];
   IF #r THEN
       "ROLL_State".M[104, 5] := TRUE;
   END_IF;
   #r := (((NOT "ROLL_State".M[190, 6]) AND "ROLL_IO".Input[5, 3] AND "ROLL_IO".Input[5, 6] AND "ROLL_IO".Input[6, 0] AND "ROLL_IO".Input[6, 2]) OR (NOT "ROLL_IO".Input[0, 1]) OR (NOT "ROLL_State".M[100, 0]) OR (NOT "ROLL_State".M[24, 1]) OR "ROLL_State".M[190, 5]);
   IF #r THEN
       "ROLL_State".M[104, 5] := FALSE;
   END_IF;
   // PB21, STEP 5 network 44
   #r := "ROLL_State".M[190, 6];
   IF #r THEN
       "ROLL_State".M[104, 6] := TRUE;
   END_IF;
   #r := (((NOT "ROLL_State".M[190, 6]) AND (("ROLL_IO".Input[5, 3] AND "ROLL_IO".Input[5, 6] AND "ROLL_IO".Input[6, 0]) OR (NOT "ROLL_IO".Input[7, 5]))) OR (NOT "ROLL_IO".Input[0, 1]) OR (NOT "ROLL_State".M[100, 0]) OR (NOT "ROLL_State".M[25, 0]) OR "ROLL_State".M[190, 5] OR "ROLL_State".M[5, 6] OR "ROLL_State".M[8, 5]);
   IF #r THEN
       "ROLL_State".M[104, 6] := FALSE;
   END_IF;
   // PB21, STEP 5 network 45
   #r := "ROLL_State".S5Timers[59].Q;
   "ROLL_IO".Output[17, 0] := #r;
   // PB21, STEP 5 network 46
   #r := ("ROLL_IO".Input[6, 5] AND "ROLL_State".M[100, 0]);
   "ROLL_IO".Output[17, 5] := #r;
   RETURN;
END_FUNCTION

FUNCTION "ROLL_PB23" : Void   // FC30, SCL
{ S7_Optimized_Access := 'TRUE' }
VERSION : 0.1
// stored: AutoNumber true, IsIECCheckEnabled false, SetENOAutomatically false, UDAEnableTagReadback false
   VAR_TEMP
      r : Bool;
      a1 : Word;
      a2 : Word;
      activeDataBlock : Int;
      comparisonResults : Array[0..0] of Bool;
   END_VAR
BEGIN

   #r := FALSE;
   #a1 := W#16#0000;
   #a2 := W#16#0000;
   #activeDataBlock := 0;
   // PB23, STEP 5 network 1
   #activeDataBlock := 15;
   // PB23, STEP 5 network 2
   #r := (("ROLL_State".M[40, 3] OR "ROLL_State".M[40, 4] OR "ROLL_State".M[40, 5]) AND "ROLL_State".M[111, 4]);
   "ROLL_State".M[240, 0] := #r;
   // PB23, STEP 5 network 3
   #a2 := #a1;
   #a1 := W#16#2120;
   #r := "ROLL_State".M[240, 0];
   "ROLL_TimerOp"(Number := 51,
                  Operation := 1,
                  Signal := #r,
                  Preset := #a1);
   #r := "ROLL_State".S5Timers[51].Q;
   "ROLL_IO".Output[19, 0] := #r;
   // PB23, STEP 5 network 4
   #a2 := #a1;
   #a1 := W#16#1050;
   #r := ((NOT "ROLL_State".M[6, 1]) AND ("ROLL_State".M[40, 4] OR "ROLL_State".M[40, 5]) AND "ROLL_IO".Output[19, 0] AND "ROLL_State".M[240, 0] AND "ROLL_State".M[35, 2] AND "ROLL_State".S5Timers[70].Q);
   "ROLL_TimerOp"(Number := 52,
                  Operation := 0,
                  Signal := #r,
                  Preset := #a1);
   #r := "ROLL_State".S5Timers[52].Q;
   "ROLL_IO".Output[19, 1] := #r;
   // PB23, STEP 5 network 5
   #r := ("ROLL_IO".Input[0, 2] AND "ROLL_IO".Input[0, 4]);
   IF #r THEN
       "ROLL_State".M[103, 7] := TRUE;
   END_IF;
   #r := (NOT "ROLL_State".S5Timers[59].Q);
   IF #r THEN
       "ROLL_State".M[103, 7] := FALSE;
   END_IF;
   // PB23, STEP 5 network 6
   #a2 := #a1;
   #a1 := W#16#3360;
   #r := "ROLL_State".S5Timers[59].Q;
   "ROLL_TimerOp"(Number := 76,
                  Operation := 0,
                  Signal := #r,
                  Preset := #a1);
   // PB23, STEP 5 network 7
   #r := ((NOT "ROLL_State".M[13, 3]) AND (NOT "ROLL_State".M[5, 6]) AND (NOT "ROLL_State".M[6, 2]) AND (NOT "ROLL_State".M[6, 3]) AND (((NOT "ROLL_State".S5Timers[76].Q) AND "ROLL_IO".Input[2, 2]) OR "ROLL_State".M[103, 7] OR "ROLL_State".M[152, 0]) AND ("ROLL_IO".Input[2, 2] OR "ROLL_State".M[152, 0]) AND "ROLL_IO".Input[3, 4] AND "ROLL_IO".Input[5, 6] AND "ROLL_State".S5Timers[59].Q);
   "ROLL_IO".Output[19, 5] := #r;
   // PB23, STEP 5 network 8
   #r := ((NOT "ROLL_State".M[5, 6]) AND (NOT "ROLL_State".M[6, 1]) AND ("ROLL_IO".Input[0, 1] OR "ROLL_IO".Input[0, 2]) AND "ROLL_IO".Input[3, 1] AND "ROLL_IO".Input[3, 4] AND "ROLL_State".M[0, 3] AND "ROLL_State".M[100, 0] AND "ROLL_State".S5Timers[70].Q);
   "ROLL_State".M[240, 0] := #r;
   // PB23, STEP 5 network 9
   #r := ((NOT "ROLL_IO".Output[20, 6]) AND (NOT "ROLL_State".M[5, 6]) AND (NOT "ROLL_State".M[8, 5]) AND (NOT "ROLL_State".S5Timers[96].Q) AND (("ROLL_State".M[100, 0] AND "ROLL_State".M[103, 1]) OR "ROLL_State".M[102, 6] OR "ROLL_State".M[104, 6]));
   "ROLL_IO".Output[20, 4] := #r;
   "ROLL_IO".Output[22, 6] := #r;
   // PB23, STEP 5 network 10
   #r := ((NOT "ROLL_IO".Output[20, 1]) AND ("ROLL_State".M[104, 0] OR "ROLL_State".M[104, 1] OR "ROLL_State".M[104, 4] OR "ROLL_State".M[152, 1]) AND "ROLL_State".M[99, 7]);
   "ROLL_IO".Output[20, 6] := #r;
   // PB23, STEP 5 network 11
   #r := ("ROLL_State".M[102, 7] OR "ROLL_State".M[103, 2] OR "ROLL_State".M[104, 5]);
   "ROLL_State".M[240, 0] := #r;
   // PB23, STEP 5 network 12
   #r := ((NOT "ROLL_State".M[13, 4]) AND (NOT "ROLL_State".M[6, 0]) AND (NOT "ROLL_State".M[6, 2]) AND (NOT "ROLL_State".M[7, 7]) AND "ROLL_IO".Input[3, 1] AND "ROLL_IO".Input[5, 0] AND "ROLL_IO".Input[5, 2] AND "ROLL_IO".Input[5, 4] AND "ROLL_State".M[240, 0]);
   "ROLL_IO".Output[20, 1] := #r;
   // PB23, STEP 5 network 13
   #r := "ROLL_State".M[103, 1];
   "ROLL_IO".Output[22, 2] := #r;
   // PB23, STEP 5 network 14
   #r := ("ROLL_State".M[102, 1] OR "ROLL_State".M[102, 2] OR "ROLL_State".M[102, 3] OR "ROLL_State".M[102, 6] OR "ROLL_State".M[102, 7] OR "ROLL_State".M[103, 2]);
   "ROLL_IO".Output[22, 3] := #r;
   // PB23, STEP 5 network 15
   #r := "ROLL_State".S5Timers[85].Q;
   "ROLL_IO".Output[21, 3] := #r;
   // PB23, STEP 5 network 16
   #a2 := #a1;
   #a1 := W#16#1020;
   #r := "ROLL_IO".Output[20, 6];
   "ROLL_TimerOp"(Number := 47,
                  Operation := 1,
                  Signal := #r,
                  Preset := #a1);
   // PB23, STEP 5 network 17
   #r := ((NOT "ROLL_IO".Output[21, 5]) AND (NOT "ROLL_IO".Output[22, 3]) AND (NOT "ROLL_IO".Output[22, 6]) AND (("ROLL_IO".Output[21, 4] AND "ROLL_State".S5Timers[47].Q) OR "ROLL_State".M[104, 0] OR "ROLL_State".M[152, 1]));
   "ROLL_IO".Output[21, 4] := #r;
   // PB23, STEP 5 network 18
   #r := ((NOT "ROLL_IO".Output[21, 4]) AND "ROLL_State".M[152, 0]);
   "ROLL_IO".Output[21, 5] := #r;
   // PB23, STEP 5 network 19
   RETURN;
END_FUNCTION

FUNCTION "ROLL_PB24" : Void   // FC31, SCL
{ S7_Optimized_Access := 'TRUE' }
VERSION : 0.1
// stored: AutoNumber true, IsIECCheckEnabled false, SetENOAutomatically false, UDAEnableTagReadback false
   VAR_TEMP
      r : Bool;
      a1 : Word;
      a2 : Word;
      activeDataBlock : Int;
      comparisonResults : Array[0..0] of Bool;
   END_VAR
BEGIN

   #r := FALSE;
   #a1 := W#16#0000;
   #a2 := W#16#0000;
   #activeDataBlock := 0;
   // PB24, STEP 5 network 1
   #activeDataBlock := 15;
   // PB24, STEP 5 network 2
   #r := ("ROLL_IO".Input[5, 0] AND "ROLL_State".M[13, 3] AND "ROLL_State".S5Timers[59].Q);
   "ROLL_State".M[240, 0] := #r;
   // PB24, STEP 5 network 3
   #a2 := #a1;
   #a1 := "ROLL_GetDW"(DbNumber := #activeDataBlock, Index := 54);
   #r := (NOT "ROLL_State".S5Timers[53].Q);
   "ROLL_TimerOp"(Number := 54,
                  Operation := 0,
                  Signal := #r,
                  Preset := #a1);
   #a2 := #a1;
   #a1 := "ROLL_GetDW"(DbNumber := #activeDataBlock, Index := 53);
   #r := "ROLL_State".S5Timers[54].Q;
   "ROLL_TimerOp"(Number := 53,
                  Operation := 1,
                  Signal := #r,
                  Preset := #a1);
   #r := "ROLL_State".M[240, 0];
   "ROLL_TimerOp"(Number := 53,
                  Operation := 2,
                  Signal := #r,
                  Preset := #a1);
   #r := ((NOT "ROLL_State".M[40, 5]) AND "ROLL_State".S5Timers[53].Q);
   "ROLL_IO".Output[19, 4] := #r;
   // PB24, STEP 5 network 4
   RETURN;
END_FUNCTION

FUNCTION "ROLL_PB25" : Void   // FC32, SCL
{ S7_Optimized_Access := 'TRUE' }
VERSION : 0.1
// stored: AutoNumber true, IsIECCheckEnabled false, SetENOAutomatically false, UDAEnableTagReadback false
   VAR_TEMP
      r : Bool;
      a1 : Word;
      a2 : Word;
      activeDataBlock : Int;
      comparisonResults : Array[0..14] of Bool;
   END_VAR
BEGIN

   #r := FALSE;
   #a1 := W#16#0000;
   #a2 := W#16#0000;
   #activeDataBlock := 0;
   // PB25, STEP 5 network 1
   #activeDataBlock := 15;
   // PB25, STEP 5 network 2
   #a2 := #a1;
   #a1 := "ROLL_GetM"(FirstByte := 5, Width := 8);
   #a2 := #a1;
   #a1 := W#16#0000;
   #comparisonResults[0] := (WORD_TO_INT(#a2) <> WORD_TO_INT(#a1));
   #r := #comparisonResults[0];
   "ROLL_State".M[87, 0] := #r;
   // PB25, STEP 5 network 3
   #a2 := #a1;
   #a1 := "ROLL_GetM"(FirstByte := 6, Width := 8);
   #a2 := #a1;
   #a1 := W#16#0000;
   #comparisonResults[1] := (WORD_TO_INT(#a2) <> WORD_TO_INT(#a1));
   #r := #comparisonResults[1];
   "ROLL_State".M[87, 1] := #r;
   // PB25, STEP 5 network 4
   #a2 := #a1;
   #a1 := "ROLL_GetM"(FirstByte := 7, Width := 8);
   #a2 := #a1;
   #a1 := W#16#0000;
   #comparisonResults[2] := (WORD_TO_INT(#a2) <> WORD_TO_INT(#a1));
   #r := #comparisonResults[2];
   "ROLL_State".M[87, 2] := #r;
   // PB25, STEP 5 network 5
   #a2 := #a1;
   #a1 := "ROLL_GetM"(FirstByte := 8, Width := 8);
   #a2 := #a1;
   #a1 := W#16#0000;
   #comparisonResults[3] := (WORD_TO_INT(#a2) <> WORD_TO_INT(#a1));
   #r := #comparisonResults[3];
   "ROLL_State".M[87, 3] := #r;
   // PB25, STEP 5 network 6
   #a2 := #a1;
   #a1 := "ROLL_GetM"(FirstByte := 9, Width := 8);
   #a2 := #a1;
   #a1 := W#16#0000;
   #comparisonResults[4] := (WORD_TO_INT(#a2) <> WORD_TO_INT(#a1));
   #r := #comparisonResults[4];
   "ROLL_State".M[87, 4] := #r;
   // PB25, STEP 5 network 7
   #a2 := #a1;
   #a1 := "ROLL_GetM"(FirstByte := 10, Width := 8);
   #a2 := #a1;
   #a1 := W#16#0000;
   #comparisonResults[5] := (WORD_TO_INT(#a2) <> WORD_TO_INT(#a1));
   #r := #comparisonResults[5];
   "ROLL_State".M[87, 5] := #r;
   // PB25, STEP 5 network 8
   #a2 := #a1;
   #a1 := "ROLL_GetM"(FirstByte := 11, Width := 8);
   #a2 := #a1;
   #a1 := W#16#0000;
   #comparisonResults[6] := (WORD_TO_INT(#a2) <> WORD_TO_INT(#a1));
   #r := #comparisonResults[6];
   "ROLL_State".M[87, 6] := #r;
   // PB25, STEP 5 network 9
   #a2 := #a1;
   #a1 := "ROLL_GetM"(FirstByte := 12, Width := 8);
   #a2 := #a1;
   #a1 := W#16#0000;
   #comparisonResults[7] := (WORD_TO_INT(#a2) <> WORD_TO_INT(#a1));
   #r := #comparisonResults[7];
   "ROLL_State".M[87, 7] := #r;
   // PB25, STEP 5 network 10
   #a2 := #a1;
   #a1 := "ROLL_GetM"(FirstByte := 13, Width := 8);
   #a2 := #a1;
   #a1 := W#16#0000;
   #comparisonResults[8] := (WORD_TO_INT(#a2) <> WORD_TO_INT(#a1));
   #r := #comparisonResults[8];
   "ROLL_State".M[88, 0] := #r;
   // PB25, STEP 5 network 11
   #a2 := #a1;
   #a1 := "ROLL_GetM"(FirstByte := 14, Width := 8);
   #a2 := #a1;
   #a1 := W#16#0000;
   #comparisonResults[9] := (WORD_TO_INT(#a2) <> WORD_TO_INT(#a1));
   #r := #comparisonResults[9];
   "ROLL_State".M[88, 1] := #r;
   // PB25, STEP 5 network 12
   #a2 := #a1;
   #a1 := "ROLL_GetM"(FirstByte := 15, Width := 8);
   #a2 := #a1;
   #a1 := W#16#0000;
   #comparisonResults[10] := (WORD_TO_INT(#a2) <> WORD_TO_INT(#a1));
   #r := #comparisonResults[10];
   "ROLL_State".M[88, 2] := #r;
   // PB25, STEP 5 network 13
   #a2 := #a1;
   #a1 := "ROLL_GetM"(FirstByte := 16, Width := 8);
   #a2 := #a1;
   #a1 := W#16#0000;
   #comparisonResults[11] := (WORD_TO_INT(#a2) <> WORD_TO_INT(#a1));
   #r := #comparisonResults[11];
   "ROLL_State".M[88, 3] := #r;
   // PB25, STEP 5 network 14
   #a2 := #a1;
   #a1 := "ROLL_GetM"(FirstByte := 17, Width := 8);
   #a2 := #a1;
   #a1 := W#16#0000;
   #comparisonResults[12] := (WORD_TO_INT(#a2) <> WORD_TO_INT(#a1));
   #r := #comparisonResults[12];
   "ROLL_State".M[88, 4] := #r;
   // PB25, STEP 5 network 15
   #a2 := #a1;
   #a1 := "ROLL_GetM"(FirstByte := 18, Width := 8);
   #a2 := #a1;
   #a1 := W#16#0000;
   #comparisonResults[13] := (WORD_TO_INT(#a2) <> WORD_TO_INT(#a1));
   #r := #comparisonResults[13];
   "ROLL_State".M[88, 5] := #r;
   // PB25, STEP 5 network 16
   #a2 := #a1;
   #a1 := "ROLL_GetM"(FirstByte := 19, Width := 8);
   #a2 := #a1;
   #a1 := W#16#0000;
   #comparisonResults[14] := (WORD_TO_INT(#a2) <> WORD_TO_INT(#a1));
   #r := #comparisonResults[14];
   "ROLL_State".M[88, 6] := #r;
   // PB25, STEP 5 network 17
   #r := ("ROLL_State".M[87, 0] OR "ROLL_State".M[87, 1] OR "ROLL_State".M[87, 2] OR "ROLL_State".M[87, 3] OR "ROLL_State".M[87, 4] OR "ROLL_State".M[87, 5] OR "ROLL_State".M[87, 6] OR "ROLL_State".M[87, 7] OR "ROLL_State".M[88, 0] OR "ROLL_State".M[88, 1] OR "ROLL_State".M[88, 2] OR "ROLL_State".M[88, 3] OR "ROLL_State".M[88, 4] OR "ROLL_State".M[88, 5] OR "ROLL_State".M[88, 6]);
   "ROLL_State".M[88, 7] := #r;
   // PB25, STEP 5 network 18
   #r := ("ROLL_IO".Input[1, 2] OR "ROLL_State".M[88, 7]);
   "ROLL_IO".Output[16, 4] := #r;
   // PB25, STEP 5 network 19
   #r := (("ROLL_State".M[3, 6] AND "ROLL_State".M[31, 6]) OR "ROLL_IO".Input[1, 2]);
   "ROLL_IO".Output[16, 5] := #r;
   // PB25, STEP 5 network 20
   #r := ("ROLL_IO".Input[1, 2] OR "ROLL_IO".Input[3, 4]);
   "ROLL_IO".Output[16, 0] := #r;
   // PB25, STEP 5 network 21
   #r := (((NOT "ROLL_State".M[31, 5]) AND "ROLL_State".M[28, 4]) OR ("ROLL_State".M[3, 6] AND "ROLL_State".M[74, 0]) OR "ROLL_IO".Input[1, 2]);
   "ROLL_IO".Output[16, 2] := #r;
   // PB25, STEP 5 network 22
   #r := (("ROLL_State".M[3, 6] AND "ROLL_State".M[31, 5]) OR "ROLL_IO".Input[1, 2] OR "ROLL_State".M[31, 4]);
   "ROLL_IO".Output[16, 3] := #r;
   // PB25, STEP 5 network 23
   #r := "ROLL_IO".Input[2, 0];
   "ROLL_IO".Output[19, 3] := #r;
   // PB25, STEP 5 network 24
   #r := (((("ROLL_IO".Input[14, 0] AND "ROLL_State".M[37, 1]) OR "ROLL_State".M[53, 6]) AND "ROLL_IO".Input[0, 2]) OR ("ROLL_IO".Input[0, 1] AND "ROLL_State".M[190, 6] AND "ROLL_State".M[20, 7]));
   IF #r THEN
       "ROLL_State".M[71, 5] := TRUE;
   END_IF;
   #r := (("ROLL_IO".Input[0, 1] AND "ROLL_State".M[190, 5] AND "ROLL_State".M[20, 7]) OR ("ROLL_IO".Input[0, 2] AND "ROLL_State".M[37, 2]));
   IF #r THEN
       "ROLL_State".M[71, 5] := FALSE;
   END_IF;
   #r := "ROLL_State".M[71, 5];
   "ROLL_IO".Output[17, 7] := #r;
   // PB25, STEP 5 network 25
   RETURN;
END_FUNCTION

FUNCTION "ROLL_PB3" : Void   // FC15, SCL
{ S7_Optimized_Access := 'TRUE' }
VERSION : 0.1
// stored: AutoNumber true, IsIECCheckEnabled false, SetENOAutomatically false, UDAEnableTagReadback false
   VAR_TEMP
      r : Bool;
      a1 : Word;
      a2 : Word;
      activeDataBlock : Int;
      comparisonResults : Array[0..15] of Bool;
   END_VAR
BEGIN

   #r := FALSE;
   #a1 := W#16#0000;
   #a2 := W#16#0000;
   #activeDataBlock := 0;
   // PB3, STEP 5 network 1
   #a2 := #a1;
   #a1 := "ROLL_GetM"(FirstByte := 239, Width := 8);
   #a2 := #a1;
   #a1 := W#16#0001;
   #comparisonResults[0] := (WORD_TO_INT(#a2) = WORD_TO_INT(#a1));
   #r := #comparisonResults[0];
   "ROLL_State".M[20, 1] := #r;
   // PB3, STEP 5 network 2
   #a2 := #a1;
   #a1 := "ROLL_GetM"(FirstByte := 239, Width := 8);
   #a2 := #a1;
   #a1 := W#16#0002;
   #comparisonResults[1] := (WORD_TO_INT(#a2) = WORD_TO_INT(#a1));
   #r := #comparisonResults[1];
   "ROLL_State".M[20, 2] := #r;
   // PB3, STEP 5 network 3
   #a2 := #a1;
   #a1 := "ROLL_GetM"(FirstByte := 239, Width := 8);
   #a2 := #a1;
   #a1 := W#16#0003;
   #comparisonResults[2] := (WORD_TO_INT(#a2) = WORD_TO_INT(#a1));
   #r := #comparisonResults[2];
   "ROLL_State".M[20, 3] := #r;
   // PB3, STEP 5 network 4
   #a2 := #a1;
   #a1 := "ROLL_GetM"(FirstByte := 239, Width := 8);
   #a2 := #a1;
   #a1 := W#16#0004;
   #comparisonResults[3] := (WORD_TO_INT(#a2) = WORD_TO_INT(#a1));
   #r := #comparisonResults[3];
   "ROLL_State".M[20, 4] := #r;
   // PB3, STEP 5 network 5
   #a2 := #a1;
   #a1 := "ROLL_GetM"(FirstByte := 239, Width := 8);
   #a2 := #a1;
   #a1 := W#16#0005;
   #comparisonResults[4] := (WORD_TO_INT(#a2) = WORD_TO_INT(#a1));
   #r := #comparisonResults[4];
   "ROLL_State".M[20, 5] := #r;
   // PB3, STEP 5 network 6
   #a2 := #a1;
   #a1 := "ROLL_GetM"(FirstByte := 239, Width := 8);
   #a2 := #a1;
   #a1 := W#16#0007;
   #comparisonResults[5] := (WORD_TO_INT(#a2) = WORD_TO_INT(#a1));
   #r := #comparisonResults[5];
   "ROLL_State".M[20, 7] := #r;
   // PB3, STEP 5 network 7
   #a2 := #a1;
   #a1 := "ROLL_GetM"(FirstByte := 239, Width := 8);
   #a2 := #a1;
   #a1 := W#16#000A;
   #comparisonResults[6] := (WORD_TO_INT(#a2) = WORD_TO_INT(#a1));
   #r := #comparisonResults[6];
   "ROLL_State".M[22, 0] := #r;
   // PB3, STEP 5 network 8
   #a2 := #a1;
   #a1 := "ROLL_GetM"(FirstByte := 239, Width := 8);
   #a2 := #a1;
   #a1 := W#16#000B;
   #comparisonResults[7] := (WORD_TO_INT(#a2) = WORD_TO_INT(#a1));
   #r := #comparisonResults[7];
   "ROLL_State".M[22, 1] := #r;
   // PB3, STEP 5 network 9
   #a2 := #a1;
   #a1 := "ROLL_GetM"(FirstByte := 239, Width := 8);
   #a2 := #a1;
   #a1 := W#16#000C;
   #comparisonResults[8] := (WORD_TO_INT(#a2) = WORD_TO_INT(#a1));
   #r := #comparisonResults[8];
   "ROLL_State".M[22, 2] := #r;
   // PB3, STEP 5 network 10
   #a2 := #a1;
   #a1 := "ROLL_GetM"(FirstByte := 239, Width := 8);
   #a2 := #a1;
   #a1 := W#16#000D;
   #comparisonResults[9] := (WORD_TO_INT(#a2) = WORD_TO_INT(#a1));
   #r := #comparisonResults[9];
   "ROLL_State".M[22, 3] := #r;
   // PB3, STEP 5 network 11
   #a2 := #a1;
   #a1 := "ROLL_GetM"(FirstByte := 239, Width := 8);
   #a2 := #a1;
   #a1 := W#16#000E;
   #comparisonResults[10] := (WORD_TO_INT(#a2) = WORD_TO_INT(#a1));
   #r := #comparisonResults[10];
   "ROLL_State".M[22, 4] := #r;
   // PB3, STEP 5 network 12
   #a2 := #a1;
   #a1 := "ROLL_GetM"(FirstByte := 239, Width := 8);
   #a2 := #a1;
   #a1 := W#16#000F;
   #comparisonResults[11] := (WORD_TO_INT(#a2) = WORD_TO_INT(#a1));
   #r := #comparisonResults[11];
   "ROLL_State".M[22, 5] := #r;
   // PB3, STEP 5 network 13
   #a2 := #a1;
   #a1 := "ROLL_GetM"(FirstByte := 239, Width := 8);
   #a2 := #a1;
   #a1 := W#16#0014;
   #comparisonResults[12] := (WORD_TO_INT(#a2) = WORD_TO_INT(#a1));
   #r := #comparisonResults[12];
   "ROLL_State".M[23, 0] := #r;
   // PB3, STEP 5 network 14
   #a2 := #a1;
   #a1 := "ROLL_GetM"(FirstByte := 239, Width := 8);
   #a2 := #a1;
   #a1 := W#16#0015;
   #comparisonResults[13] := (WORD_TO_INT(#a2) = WORD_TO_INT(#a1));
   #r := #comparisonResults[13];
   "ROLL_State".M[23, 1] := #r;
   // PB3, STEP 5 network 15
   #a2 := #a1;
   #a1 := "ROLL_GetM"(FirstByte := 239, Width := 8);
   #a2 := #a1;
   #a1 := W#16#0016;
   #comparisonResults[14] := (WORD_TO_INT(#a2) = WORD_TO_INT(#a1));
   #r := #comparisonResults[14];
   "ROLL_State".M[23, 2] := #r;
   // PB3, STEP 5 network 16
   #a2 := #a1;
   #a1 := "ROLL_GetM"(FirstByte := 239, Width := 8);
   #a2 := #a1;
   #a1 := W#16#0017;
   #comparisonResults[15] := (WORD_TO_INT(#a2) = WORD_TO_INT(#a1));
   #r := #comparisonResults[15];
   "ROLL_State".M[23, 3] := #r;
   // PB3, STEP 5 network 17
   RETURN;
END_FUNCTION

FUNCTION "ROLL_PB4" : Void   // FC16, SCL
{ S7_Optimized_Access := 'TRUE' }
VERSION : 0.1
// stored: AutoNumber true, IsIECCheckEnabled false, SetENOAutomatically false, UDAEnableTagReadback false
   VAR_TEMP
      r : Bool;
      a1 : Word;
      a2 : Word;
      activeDataBlock : Int;
      comparisonResults : Array[0..24] of Bool;
   END_VAR
BEGIN

